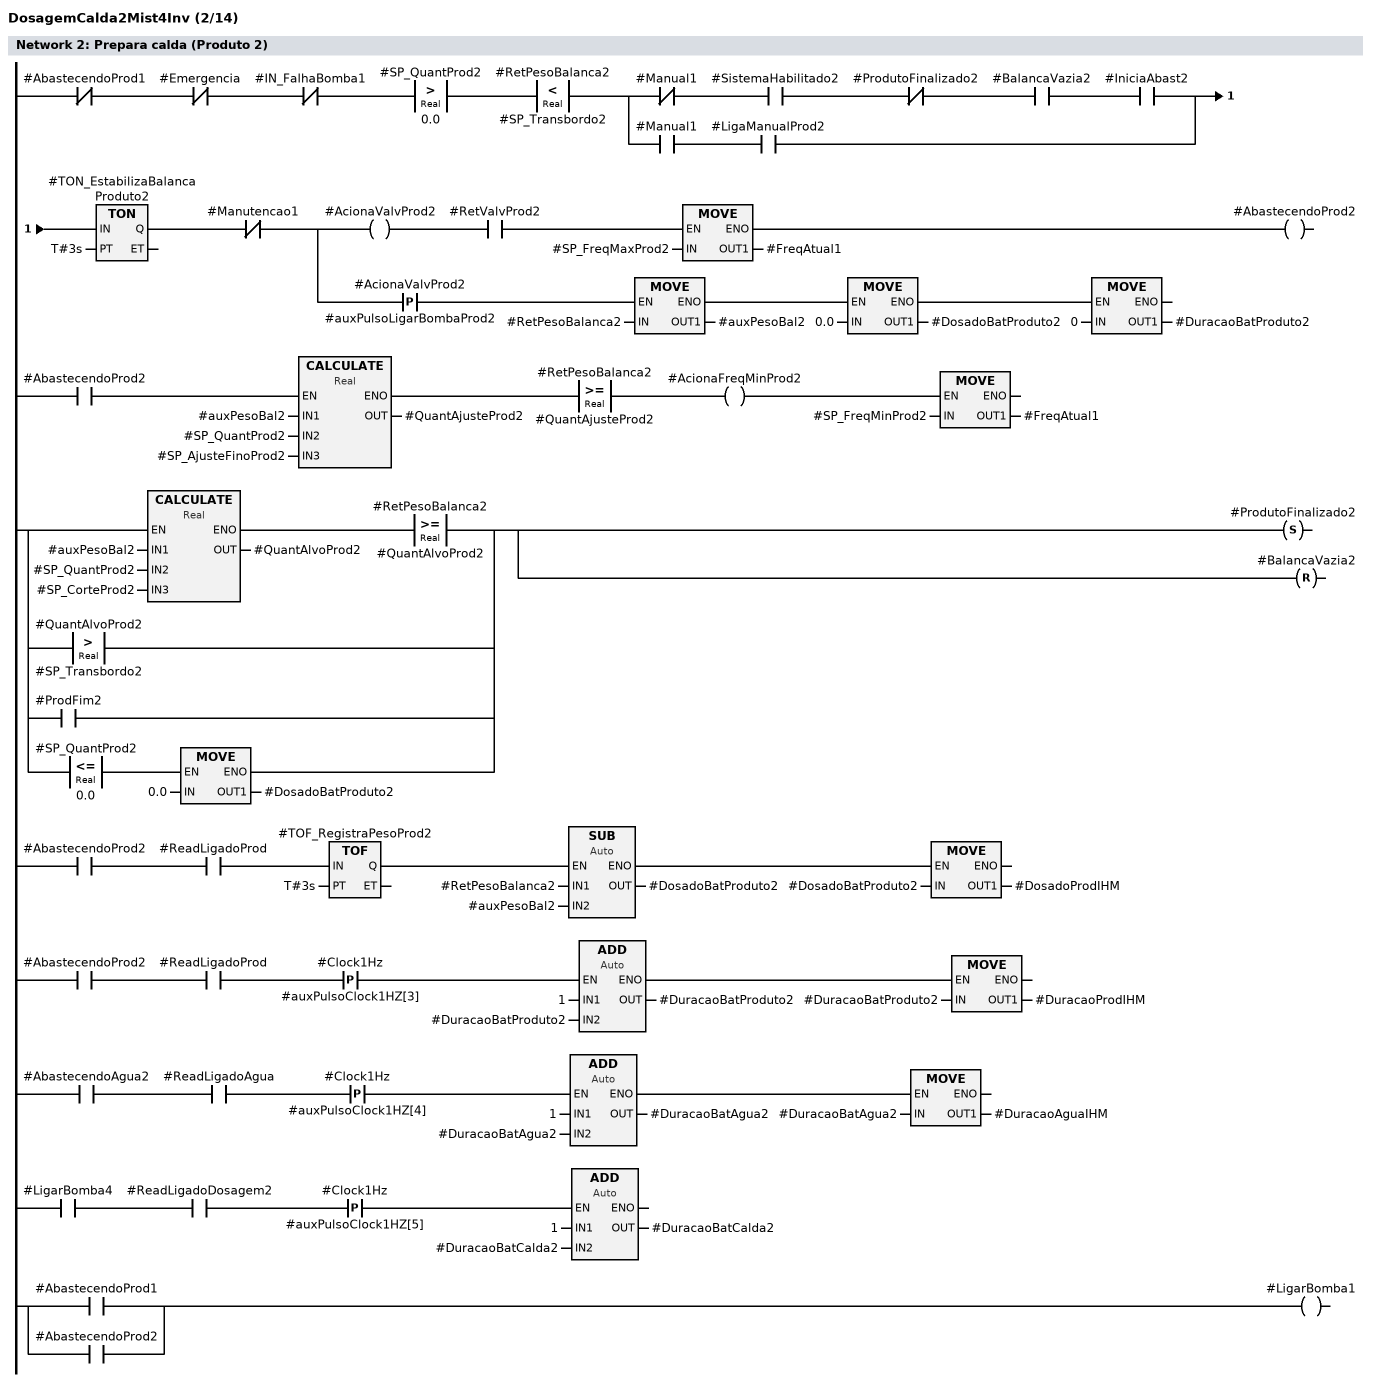
   #TON_EstabilizaBalancaProduto2(IN := NOT #AbastecendoProd1 AND NOT #Emergencia AND NOT #IN_FalhaBomba1 AND (#SP_QuantProd2 > 0.0) AND (#RetPesoBalanca2 < #SP_Transbordo2) AND ((NOT #Manual1 AND #SistemaHabilitado2 AND NOT #ProdutoFinalizado2 AND #BalancaVazia2 AND #IniciaAbast2) OR (#Manual1 AND #LigaManualProd2)),   // TON
                           PT := T#3s);
   #AcionaValvProd2 := #TON_EstabilizaBalancaProduto2.Q AND NOT #Manutencao1;
   #_w1 := #AcionaValvProd2 AND #RetValvProd2;
   IF #_w1 THEN #FreqAtual1 := #SP_FreqMaxProd2; END_IF;
   #AbastecendoProd2 := #_w1;
   #_w2 := #AcionaValvProd2 AND #AcionaValvProd2 AND NOT #auxPulsoLigarBombaProd2;   // rising edge of #AcionaValvProd2
   #auxPulsoLigarBombaProd2 := #AcionaValvProd2;
   IF #_w2 THEN
       #auxPesoBal2 := #RetPesoBalanca2;
       #DosadoBatProduto2 := 0.0;
       #DuracaoBatProduto2 := 0;
   END_IF;
   IF #AbastecendoProd2 THEN
       #QuantAjusteProd2 := (#auxPesoBal2 + #SP_QuantProd2 - #SP_AjusteFinoProd2);
   END_IF;
   #AcionaFreqMinProd2 := #AbastecendoProd2 AND (#RetPesoBalanca2 >= #QuantAjusteProd2);
   IF #AcionaFreqMinProd2 THEN #FreqAtual1 := #SP_FreqMinProd2; END_IF;
   #QuantAlvoProd2 := (#auxPesoBal2 + #SP_QuantProd2 - #SP_CorteProd2);
   #_w3 := #SP_QuantProd2 <= 0.0;
   IF #_w3 THEN #DosadoBatProduto2 := 0.0; END_IF;
   IF (#RetPesoBalanca2 >= #QuantAlvoProd2) OR (#QuantAlvoProd2 > #SP_Transbordo2) OR #ProdFim2 OR #_w3 THEN
       #ProdutoFinalizado2 := TRUE;
       #BalancaVazia2 := FALSE;
   END_IF;
   #TOF_RegistraPesoProd2(IN := #AbastecendoProd2 AND #ReadLigadoProd, PT := T#3s);   // TOF
   IF #TOF_RegistraPesoProd2.Q THEN
       #DosadoBatProduto2 := #RetPesoBalanca2 - #auxPesoBal2;
       #DosadoProdIHM := #DosadoBatProduto2;
   END_IF;
   #_w4 := #AbastecendoProd2 AND #ReadLigadoProd AND #Clock1Hz AND NOT #auxPulsoClock1HZ[3];   // rising edge of #Clock1Hz
   #auxPulsoClock1HZ[3] := #Clock1Hz;
   IF #_w4 THEN
       #DuracaoBatProduto2 := 1 + #DuracaoBatProduto2;
       #DuracaoProdIHM := #DuracaoBatProduto2;
   END_IF;
   #_w5 := #AbastecendoAgua2 AND #ReadLigadoAgua AND #Clock1Hz AND NOT #auxPulsoClock1HZ[4];   // rising edge of #Clock1Hz
   #auxPulsoClock1HZ[4] := #Clock1Hz;
   IF #_w5 THEN
       #DuracaoBatAgua2 := 1 + #DuracaoBatAgua2;
       #DuracaoAguaIHM := #DuracaoBatAgua2;
   END_IF;
   #_w6 := #LigarBomba4 AND #ReadLigadoDosagem2 AND #Clock1Hz AND NOT #auxPulsoClock1HZ[5];   // rising edge of #Clock1Hz
   #auxPulsoClock1HZ[5] := #Clock1Hz;
   IF #_w6 THEN #DuracaoBatCalda2 := 1 + #DuracaoBatCalda2; END_IF;
   #LigarBomba1 := #AbastecendoProd1 OR #AbastecendoProd2;
END_REGION

REGION Network 3: Prepara calda (Agua 1)
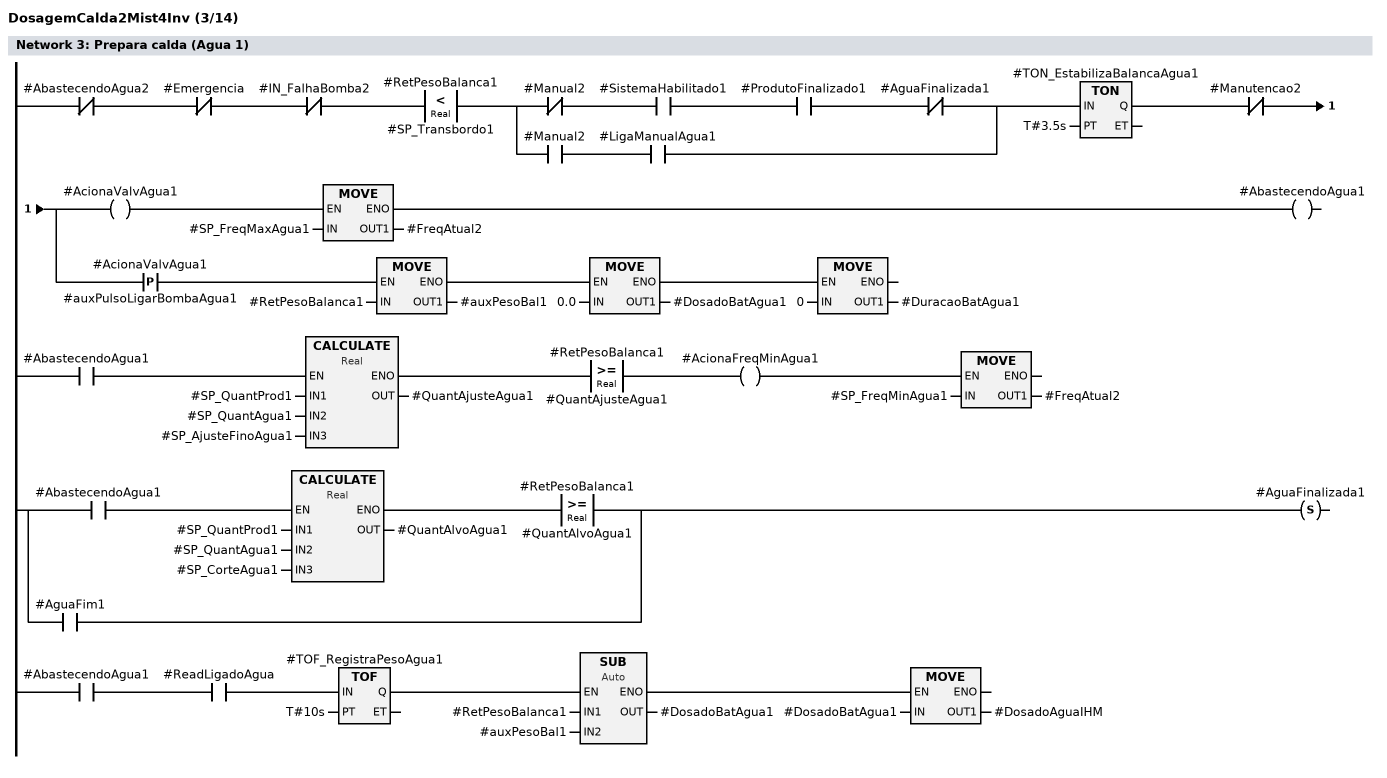
   #TON_EstabilizaBalancaAgua1(IN := NOT #AbastecendoAgua2 AND NOT #Emergencia AND NOT #IN_FalhaBomba2 AND (#RetPesoBalanca1 < #SP_Transbordo1) AND ((NOT #Manual2 AND #SistemaHabilitado1 AND #ProdutoFinalizado1 AND NOT #AguaFinalizada1) OR (#Manual2 AND #LigaManualAgua1)),   // TON
                           PT := T#3.5s);
   #AcionaValvAgua1 := #TON_EstabilizaBalancaAgua1.Q AND NOT #Manutencao2;
   IF #AcionaValvAgua1 THEN #FreqAtual2 := #SP_FreqMaxAgua1; END_IF;
   #AbastecendoAgua1 := #AcionaValvAgua1;
   #_w1 := #AcionaValvAgua1 AND #AcionaValvAgua1 AND NOT #auxPulsoLigarBombaAgua1;   // rising edge of #AcionaValvAgua1
   #auxPulsoLigarBombaAgua1 := #AcionaValvAgua1;
   IF #_w1 THEN
       #auxPesoBal1 := #RetPesoBalanca1;
       #DosadoBatAgua1 := 0.0;
       #DuracaoBatAgua1 := 0;
   END_IF;
   IF #AbastecendoAgua1 THEN
       #QuantAjusteAgua1 := (#SP_QuantProd1 + #SP_QuantAgua1 - #SP_AjusteFinoAgua1);
   END_IF;
   #AcionaFreqMinAgua1 := #AbastecendoAgua1 AND (#RetPesoBalanca1 >= #QuantAjusteAgua1);
   IF #AcionaFreqMinAgua1 THEN #FreqAtual2 := #SP_FreqMinAgua1; END_IF;
   IF #AbastecendoAgua1 THEN #QuantAlvoAgua1 := (#SP_QuantProd1 + #SP_QuantAgua1 - #SP_CorteAgua1); END_IF;
   IF (#AbastecendoAgua1 AND (#RetPesoBalanca1 >= #QuantAlvoAgua1)) OR #AguaFim1 THEN
       #AguaFinalizada1 := TRUE;
   END_IF;
   #TOF_RegistraPesoAgua1(IN := #AbastecendoAgua1 AND #ReadLigadoAgua, PT := T#10s);   // TOF
   IF #TOF_RegistraPesoAgua1.Q THEN
       #DosadoBatAgua1 := #RetPesoBalanca1 - #auxPesoBal1;
       #DosadoAguaIHM := #DosadoBatAgua1;
   END_IF;
END_REGION

REGION Network 4: Prepara calda (Agua 2)
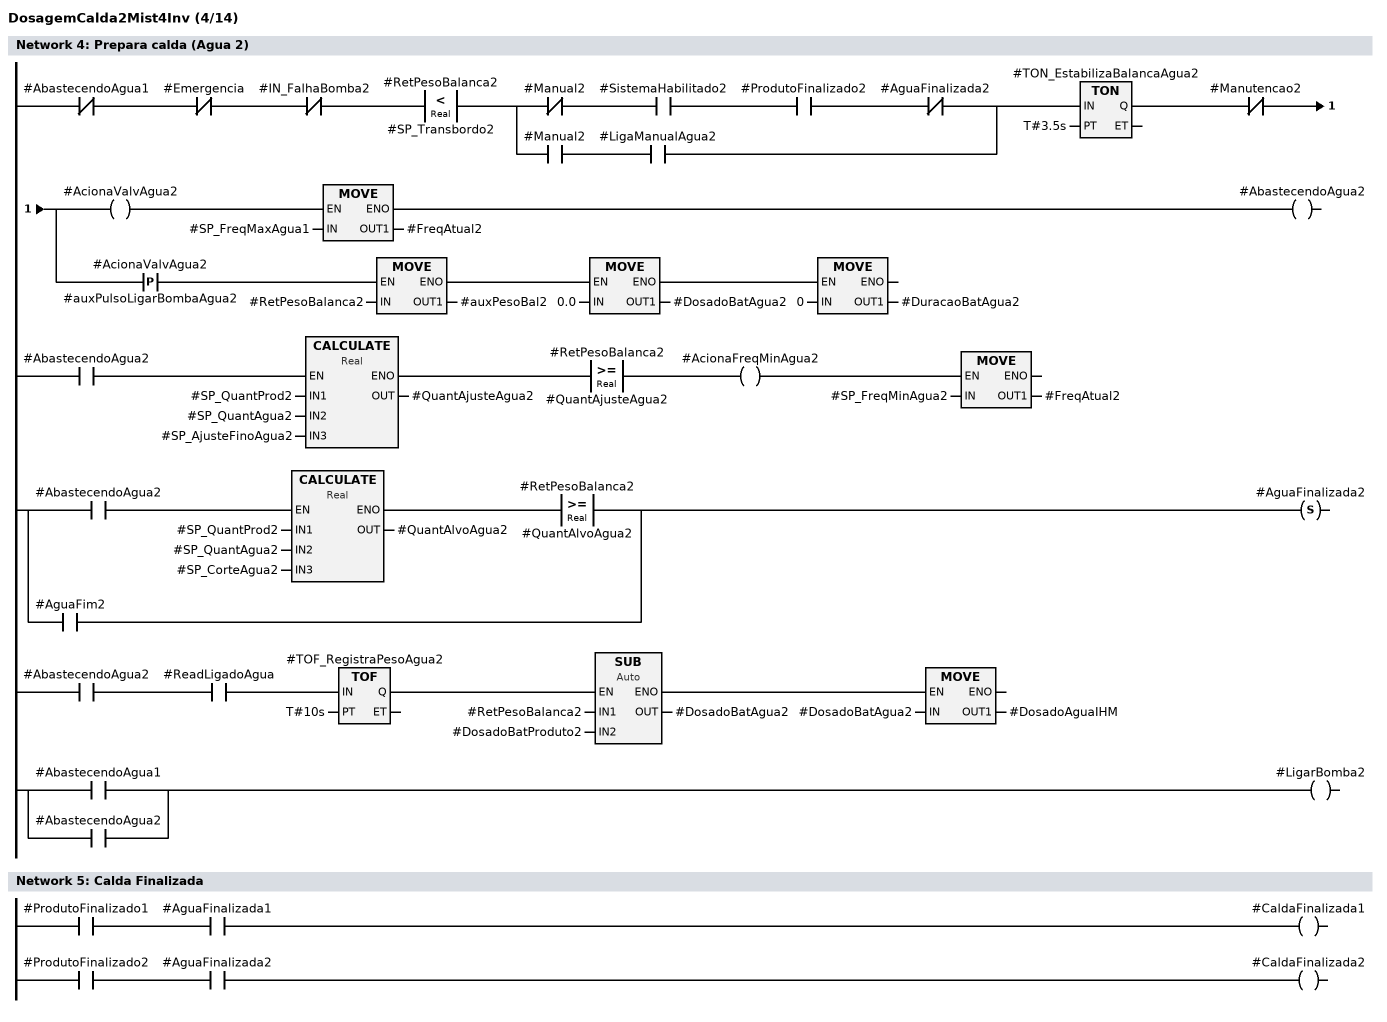
   #TON_EstabilizaBalancaAgua2(IN := NOT #AbastecendoAgua1 AND NOT #Emergencia AND NOT #IN_FalhaBomba2 AND (#RetPesoBalanca2 < #SP_Transbordo2) AND ((NOT #Manual2 AND #SistemaHabilitado2 AND #ProdutoFinalizado2 AND NOT #AguaFinalizada2) OR (#Manual2 AND #LigaManualAgua2)),   // TON
                           PT := T#3.5s);
   #AcionaValvAgua2 := #TON_EstabilizaBalancaAgua2.Q AND NOT #Manutencao2;
   IF #AcionaValvAgua2 THEN #FreqAtual2 := #SP_FreqMaxAgua1; END_IF;
   #AbastecendoAgua2 := #AcionaValvAgua2;
   #_w1 := #AcionaValvAgua2 AND #AcionaValvAgua2 AND NOT #auxPulsoLigarBombaAgua2;   // rising edge of #AcionaValvAgua2
   #auxPulsoLigarBombaAgua2 := #AcionaValvAgua2;
   IF #_w1 THEN
       #auxPesoBal2 := #RetPesoBalanca2;
       #DosadoBatAgua2 := 0.0;
       #DuracaoBatAgua2 := 0;
   END_IF;
   IF #AbastecendoAgua2 THEN
       #QuantAjusteAgua2 := (#SP_QuantProd2 + #SP_QuantAgua2 - #SP_AjusteFinoAgua2);
   END_IF;
   #AcionaFreqMinAgua2 := #AbastecendoAgua2 AND (#RetPesoBalanca2 >= #QuantAjusteAgua2);
   IF #AcionaFreqMinAgua2 THEN #FreqAtual2 := #SP_FreqMinAgua2; END_IF;
   IF #AbastecendoAgua2 THEN #QuantAlvoAgua2 := (#SP_QuantProd2 + #SP_QuantAgua2 - #SP_CorteAgua2); END_IF;
   IF (#AbastecendoAgua2 AND (#RetPesoBalanca2 >= #QuantAlvoAgua2)) OR #AguaFim2 THEN
       #AguaFinalizada2 := TRUE;
   END_IF;
   #TOF_RegistraPesoAgua2(IN := #AbastecendoAgua2 AND #ReadLigadoAgua, PT := T#10s);   // TOF
   IF #TOF_RegistraPesoAgua2.Q THEN
       #DosadoBatAgua2 := #RetPesoBalanca2 - #DosadoBatProduto2;
       #DosadoAguaIHM := #DosadoBatAgua2;
   END_IF;
   #LigarBomba2 := #AbastecendoAgua1 OR #AbastecendoAgua2;
END_REGION

REGION Network 5: Calda Finalizada
   RUNG wire#powerrail
      Contact( #ProdutoFinalizado1 )
      Contact( #AguaFinalizada1 )
      Coil( #CaldaFinalizada1 )
   END_RUNG
   RUNG wire#powerrail
      Contact( #ProdutoFinalizado2 )
      Contact( #AguaFinalizada2 )
      Coil( #CaldaFinalizada2 )
   END_RUNG
   // the same network as SCL:
   #CaldaFinalizada1 := #ProdutoFinalizado1 AND #AguaFinalizada1;
   #CaldaFinalizada2 := #ProdutoFinalizado2 AND #AguaFinalizada2;
END_REGION

REGION Network 6: Tempo de mistura seca 1
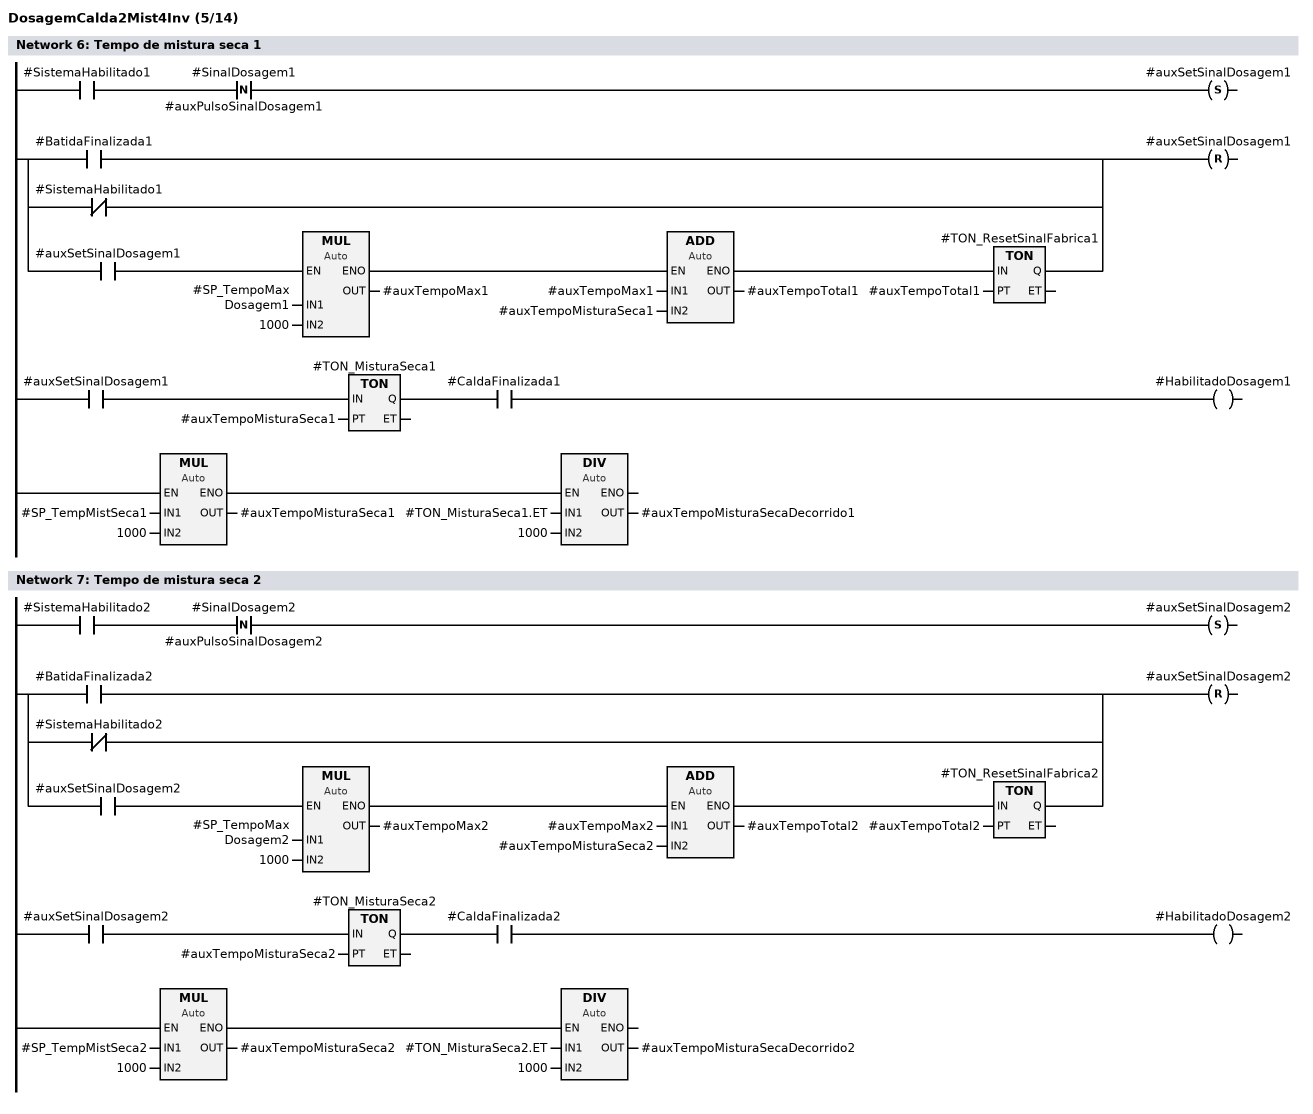
   #_w1 := #SistemaHabilitado1 AND NOT #SinalDosagem1 AND #auxPulsoSinalDosagem1;   // falling edge of #SinalDosagem1
   #auxPulsoSinalDosagem1 := #SinalDosagem1;
   IF #_w1 THEN #auxSetSinalDosagem1 := TRUE; END_IF;
   IF #auxSetSinalDosagem1 THEN
       #auxTempoMax1 := #SP_TempoMaxDosagem1 * 1000;
       #auxTempoTotal1 := #auxTempoMax1 + #auxTempoMisturaSeca1;
   END_IF;
   #TON_ResetSinalFabrica1(IN := #auxSetSinalDosagem1, PT := #auxTempoTotal1);   // TON
   IF #BatidaFinalizada1 OR NOT #SistemaHabilitado1 OR #TON_ResetSinalFabrica1.Q THEN
       #auxSetSinalDosagem1 := FALSE;
   END_IF;
   #TON_MisturaSeca1(IN := #auxSetSinalDosagem1, PT := #auxTempoMisturaSeca1);   // TON
   #HabilitadoDosagem1 := #TON_MisturaSeca1.Q AND #CaldaFinalizada1;
   #auxTempoMisturaSeca1 := #SP_TempMistSeca1 * 1000;
   #auxTempoMisturaSecaDecorrido1 := #TON_MisturaSeca1.ET / 1000;
END_REGION

REGION Network 7: Tempo de mistura seca 2
   #_w1 := #SistemaHabilitado2 AND NOT #SinalDosagem2 AND #auxPulsoSinalDosagem2;   // falling edge of #SinalDosagem2
   #auxPulsoSinalDosagem2 := #SinalDosagem2;
   IF #_w1 THEN #auxSetSinalDosagem2 := TRUE; END_IF;
   IF #auxSetSinalDosagem2 THEN
       #auxTempoMax2 := #SP_TempoMaxDosagem2 * 1000;
       #auxTempoTotal2 := #auxTempoMax2 + #auxTempoMisturaSeca2;
   END_IF;
   #TON_ResetSinalFabrica2(IN := #auxSetSinalDosagem2, PT := #auxTempoTotal2);   // TON
   IF #BatidaFinalizada2 OR NOT #SistemaHabilitado2 OR #TON_ResetSinalFabrica2.Q THEN
       #auxSetSinalDosagem2 := FALSE;
   END_IF;
   #TON_MisturaSeca2(IN := #auxSetSinalDosagem2, PT := #auxTempoMisturaSeca2);   // TON
   #HabilitadoDosagem2 := #TON_MisturaSeca2.Q AND #CaldaFinalizada2;
   #auxTempoMisturaSeca2 := #SP_TempMistSeca2 * 1000;
   #auxTempoMisturaSecaDecorrido2 := #TON_MisturaSeca2.ET / 1000;
END_REGION

REGION Network 8: Dosa calda 1
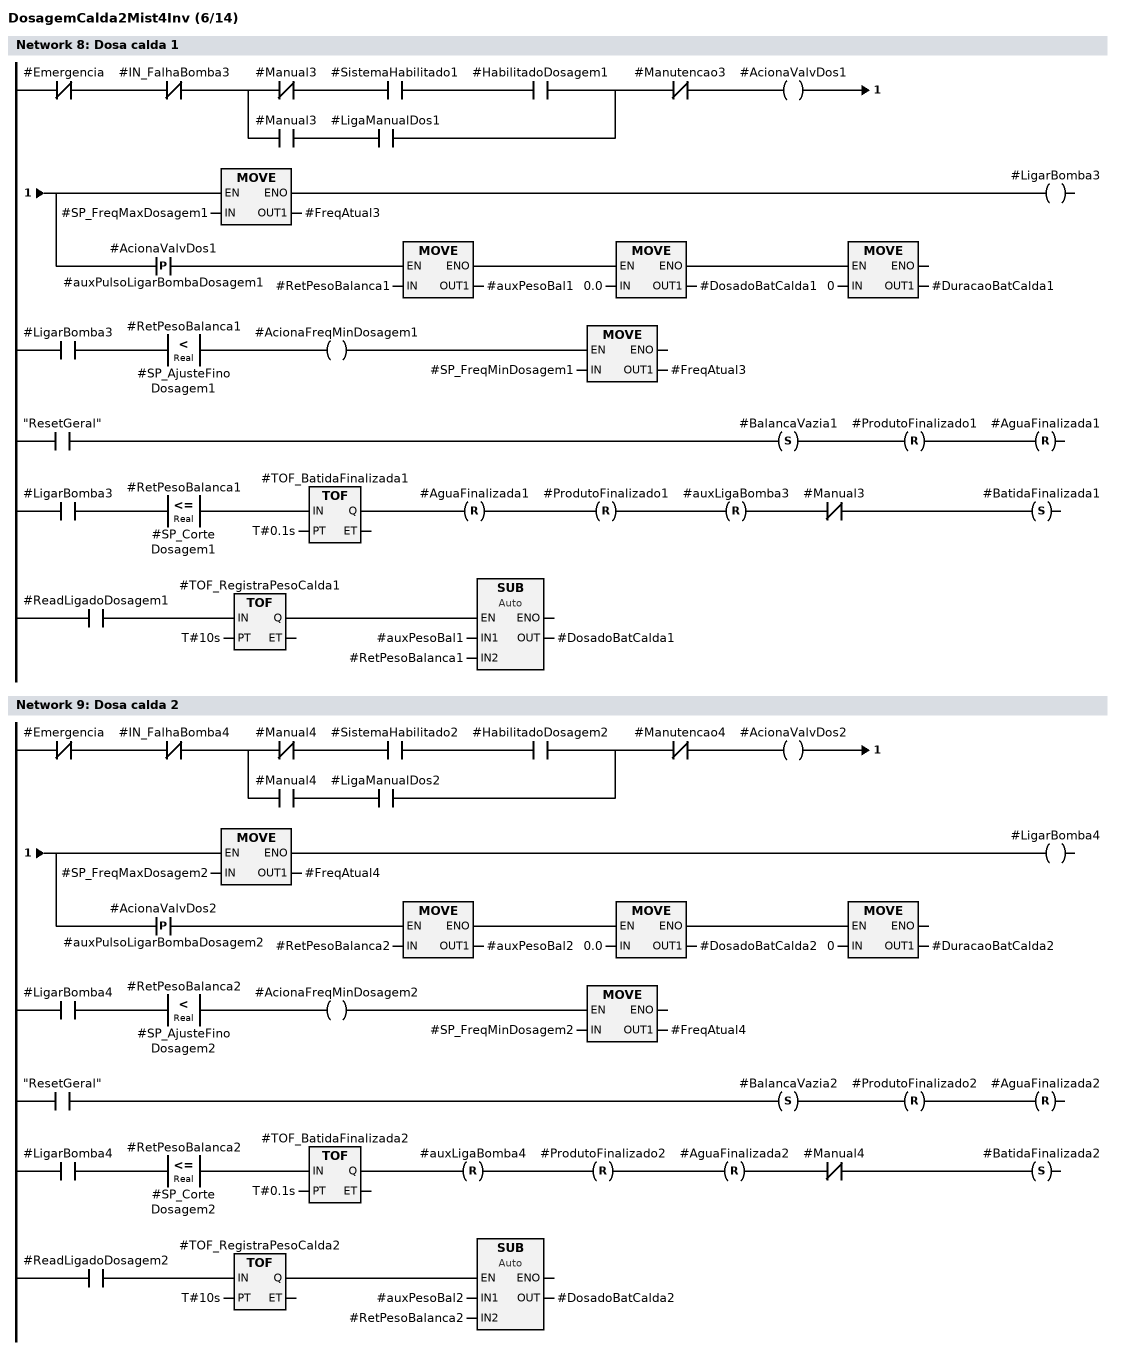
   #AcionaValvDos1 := NOT #Emergencia AND NOT #IN_FalhaBomba3 AND ((NOT #Manual3 AND #SistemaHabilitado1 AND #HabilitadoDosagem1) OR (#Manual3 AND #LigaManualDos1)) AND NOT #Manutencao3;
   IF #AcionaValvDos1 THEN #FreqAtual3 := #SP_FreqMaxDosagem1; END_IF;
   #LigarBomba3 := #AcionaValvDos1;
   #_w1 := #AcionaValvDos1 AND #AcionaValvDos1 AND NOT #auxPulsoLigarBombaDosagem1;   // rising edge of #AcionaValvDos1
   #auxPulsoLigarBombaDosagem1 := #AcionaValvDos1;
   IF #_w1 THEN
       #auxPesoBal1 := #RetPesoBalanca1;
       #DosadoBatCalda1 := 0.0;
       #DuracaoBatCalda1 := 0;
   END_IF;
   #AcionaFreqMinDosagem1 := #LigarBomba3 AND (#RetPesoBalanca1 < #SP_AjusteFinoDosagem1);
   IF #AcionaFreqMinDosagem1 THEN #FreqAtual3 := #SP_FreqMinDosagem1; END_IF;
   IF "ResetGeral" THEN
       #BalancaVazia1 := TRUE;
       #ProdutoFinalizado1 := FALSE;
       #AguaFinalizada1 := FALSE;
   END_IF;
   #TOF_BatidaFinalizada1(IN := #LigarBomba3 AND (#RetPesoBalanca1 <= #SP_CorteDosagem1), PT := T#0.1s);   // TOF
   IF #TOF_BatidaFinalizada1.Q THEN
       #AguaFinalizada1 := FALSE;
       #ProdutoFinalizado1 := FALSE;
       #auxLigaBomba3 := FALSE;
   END_IF;
   IF #TOF_BatidaFinalizada1.Q AND NOT #Manual3 THEN #BatidaFinalizada1 := TRUE; END_IF;
   #TOF_RegistraPesoCalda1(IN := #ReadLigadoDosagem1, PT := T#10s);   // TOF
   IF #TOF_RegistraPesoCalda1.Q THEN #DosadoBatCalda1 := #auxPesoBal1 - #RetPesoBalanca1; END_IF;
END_REGION

REGION Network 9: Dosa calda 2
   #AcionaValvDos2 := NOT #Emergencia AND NOT #IN_FalhaBomba4 AND ((NOT #Manual4 AND #SistemaHabilitado2 AND #HabilitadoDosagem2) OR (#Manual4 AND #LigaManualDos2)) AND NOT #Manutencao4;
   IF #AcionaValvDos2 THEN #FreqAtual4 := #SP_FreqMaxDosagem2; END_IF;
   #LigarBomba4 := #AcionaValvDos2;
   #_w1 := #AcionaValvDos2 AND #AcionaValvDos2 AND NOT #auxPulsoLigarBombaDosagem2;   // rising edge of #AcionaValvDos2
   #auxPulsoLigarBombaDosagem2 := #AcionaValvDos2;
   IF #_w1 THEN
       #auxPesoBal2 := #RetPesoBalanca2;
       #DosadoBatCalda2 := 0.0;
       #DuracaoBatCalda2 := 0;
   END_IF;
   #AcionaFreqMinDosagem2 := #LigarBomba4 AND (#RetPesoBalanca2 < #SP_AjusteFinoDosagem2);
   IF #AcionaFreqMinDosagem2 THEN #FreqAtual4 := #SP_FreqMinDosagem2; END_IF;
   IF "ResetGeral" THEN
       #BalancaVazia2 := TRUE;
       #ProdutoFinalizado2 := FALSE;
       #AguaFinalizada2 := FALSE;
   END_IF;
   #TOF_BatidaFinalizada2(IN := #LigarBomba4 AND (#RetPesoBalanca2 <= #SP_CorteDosagem2), PT := T#0.1s);   // TOF
   IF #TOF_BatidaFinalizada2.Q THEN
       #auxLigaBomba4 := FALSE;
       #ProdutoFinalizado2 := FALSE;
       #AguaFinalizada2 := FALSE;
   END_IF;
   IF #TOF_BatidaFinalizada2.Q AND NOT #Manual4 THEN #BatidaFinalizada2 := TRUE; END_IF;
   #TOF_RegistraPesoCalda2(IN := #ReadLigadoDosagem2, PT := T#10s);   // TOF
   IF #TOF_RegistraPesoCalda2.Q THEN #DosadoBatCalda2 := #auxPesoBal2 - #RetPesoBalanca2; END_IF;
END_REGION

REGION Network 10: Grava batelada
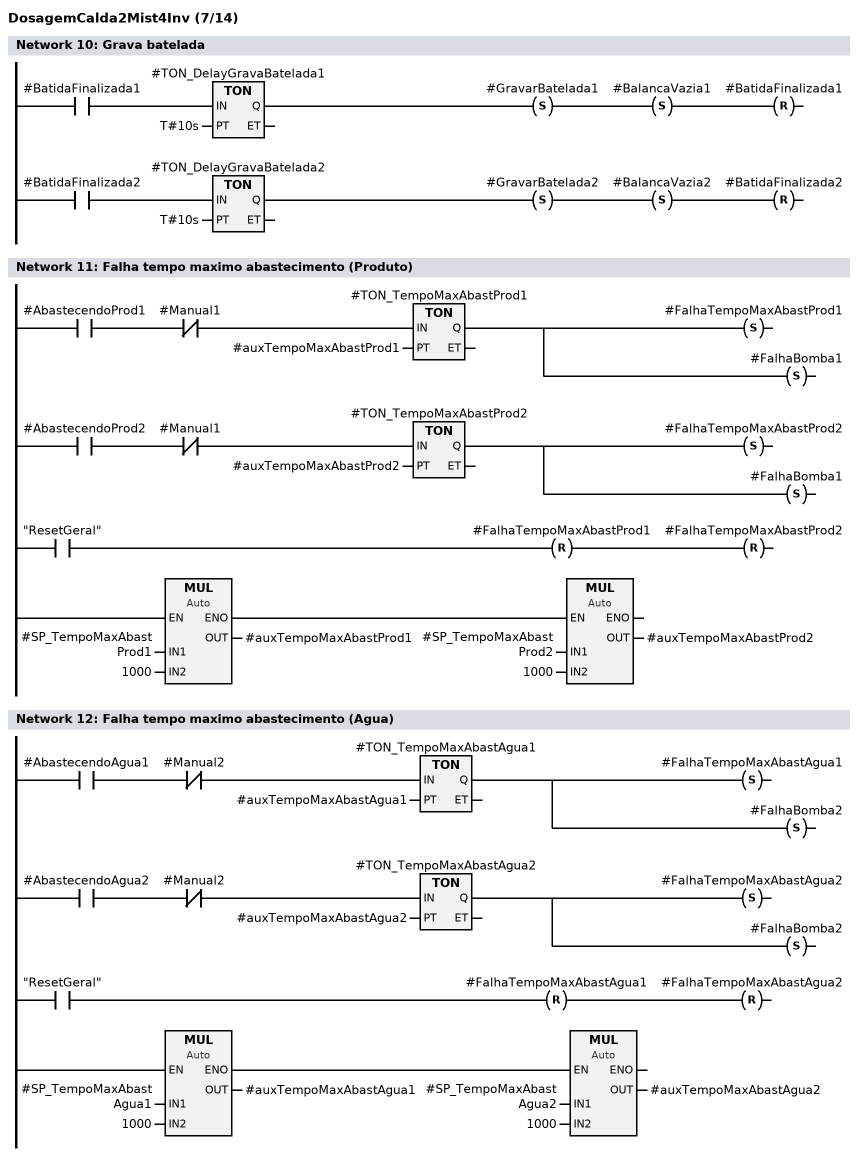
   #TON_DelayGravaBatelada1(IN := #BatidaFinalizada1, PT := T#10s);   // TON
   IF #TON_DelayGravaBatelada1.Q THEN
       #GravarBatelada1 := TRUE;
       #BalancaVazia1 := TRUE;
       #BatidaFinalizada1 := FALSE;
   END_IF;
   #TON_DelayGravaBatelada2(IN := #BatidaFinalizada2, PT := T#10s);   // TON
   IF #TON_DelayGravaBatelada2.Q THEN
       #GravarBatelada2 := TRUE;
       #BalancaVazia2 := TRUE;
       #BatidaFinalizada2 := FALSE;
   END_IF;
END_REGION

REGION Network 11: Falha tempo maximo abastecimento (Produto)
   #TON_TempoMaxAbastProd1(IN := #AbastecendoProd1 AND NOT #Manual1, PT := #auxTempoMaxAbastProd1);   // TON
   IF #TON_TempoMaxAbastProd1.Q THEN
       #FalhaTempoMaxAbastProd1 := TRUE;
       #FalhaBomba1 := TRUE;
   END_IF;
   #TON_TempoMaxAbastProd2(IN := #AbastecendoProd2 AND NOT #Manual1, PT := #auxTempoMaxAbastProd2);   // TON
   IF #TON_TempoMaxAbastProd2.Q THEN
       #FalhaTempoMaxAbastProd2 := TRUE;
       #FalhaBomba1 := TRUE;
   END_IF;
   IF "ResetGeral" THEN
       #FalhaTempoMaxAbastProd1 := FALSE;
       #FalhaTempoMaxAbastProd2 := FALSE;
   END_IF;
   #auxTempoMaxAbastProd1 := #SP_TempoMaxAbastProd1 * 1000;
   #auxTempoMaxAbastProd2 := #SP_TempoMaxAbastProd2 * 1000;
END_REGION

REGION Network 12: Falha tempo maximo abastecimento (Agua)
   #TON_TempoMaxAbastAgua1(IN := #AbastecendoAgua1 AND NOT #Manual2, PT := #auxTempoMaxAbastAgua1);   // TON
   IF #TON_TempoMaxAbastAgua1.Q THEN
       #FalhaTempoMaxAbastAgua1 := TRUE;
       #FalhaBomba2 := TRUE;
   END_IF;
   #TON_TempoMaxAbastAgua2(IN := #AbastecendoAgua2 AND NOT #Manual2, PT := #auxTempoMaxAbastAgua2);   // TON
   IF #TON_TempoMaxAbastAgua2.Q THEN
       #FalhaTempoMaxAbastAgua2 := TRUE;
       #FalhaBomba2 := TRUE;
   END_IF;
   IF "ResetGeral" THEN
       #FalhaTempoMaxAbastAgua1 := FALSE;
       #FalhaTempoMaxAbastAgua2 := FALSE;
   END_IF;
   #auxTempoMaxAbastAgua1 := #SP_TempoMaxAbastAgua1 * 1000;
   #auxTempoMaxAbastAgua2 := #SP_TempoMaxAbastAgua2 * 1000;
END_REGION

REGION Network 13: Falha tempo maximo de dosagem (Calda)
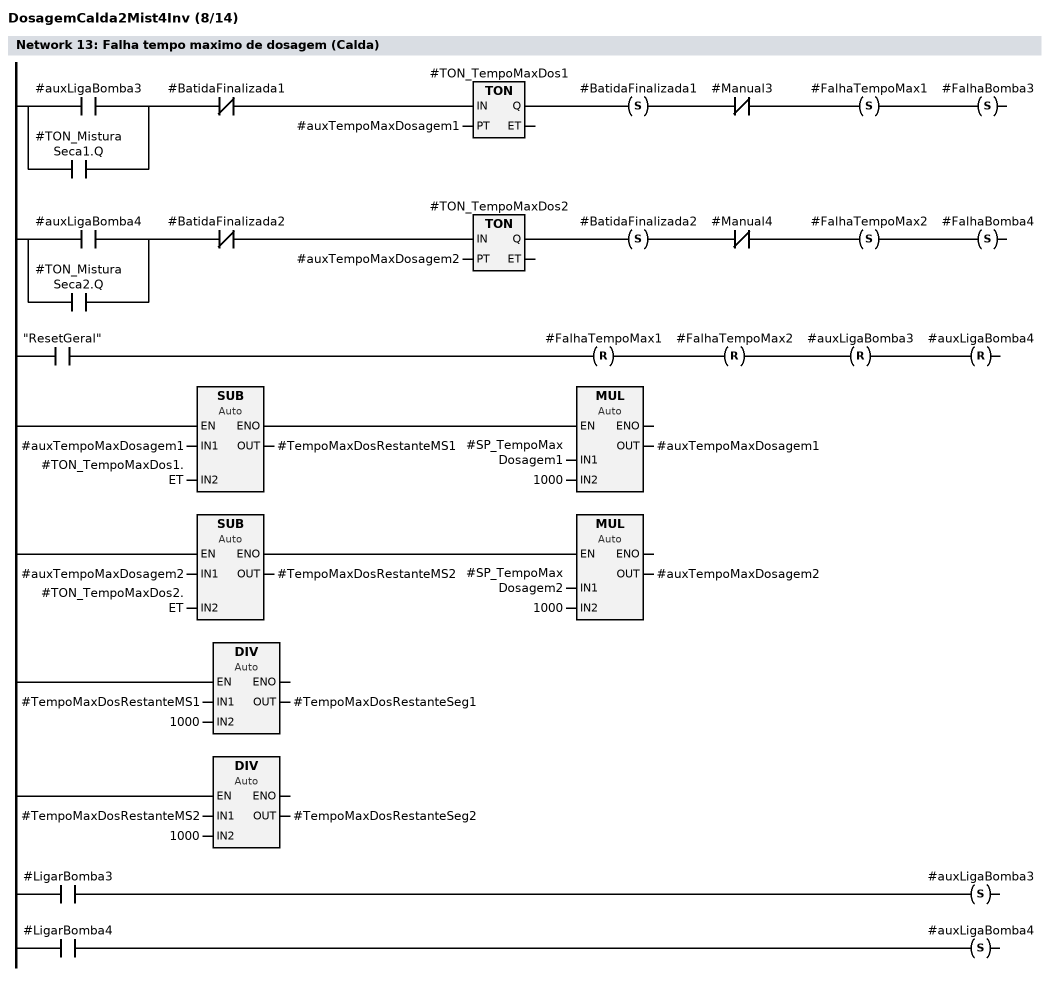
   #TON_TempoMaxDos1(IN := (#auxLigaBomba3 OR #TON_MisturaSeca1.Q) AND NOT #BatidaFinalizada1,   // TON
                     PT := #auxTempoMaxDosagem1);
   IF #TON_TempoMaxDos1.Q THEN #BatidaFinalizada1 := TRUE; END_IF;
   IF #TON_TempoMaxDos1.Q AND NOT #Manual3 THEN
       #FalhaTempoMax1 := TRUE;
       #FalhaBomba3 := TRUE;
   END_IF;
   #TON_TempoMaxDos2(IN := (#auxLigaBomba4 OR #TON_MisturaSeca2.Q) AND NOT #BatidaFinalizada2,   // TON
                     PT := #auxTempoMaxDosagem2);
   IF #TON_TempoMaxDos2.Q THEN #BatidaFinalizada2 := TRUE; END_IF;
   IF #TON_TempoMaxDos2.Q AND NOT #Manual4 THEN
       #FalhaTempoMax2 := TRUE;
       #FalhaBomba4 := TRUE;
   END_IF;
   IF "ResetGeral" THEN
       #FalhaTempoMax1 := FALSE;
       #FalhaTempoMax2 := FALSE;
       #auxLigaBomba3 := FALSE;
       #auxLigaBomba4 := FALSE;
   END_IF;
   #TempoMaxDosRestanteMS1 := #auxTempoMaxDosagem1 - #TON_TempoMaxDos1.ET;
   #auxTempoMaxDosagem1 := #SP_TempoMaxDosagem1 * 1000;
   #TempoMaxDosRestanteMS2 := #auxTempoMaxDosagem2 - #TON_TempoMaxDos2.ET;
   #auxTempoMaxDosagem2 := #SP_TempoMaxDosagem2 * 1000;
   #TempoMaxDosRestanteSeg1 := #TempoMaxDosRestanteMS1 / 1000;
   #TempoMaxDosRestanteSeg2 := #TempoMaxDosRestanteMS2 / 1000;
   IF #LigarBomba3 THEN #auxLigaBomba3 := TRUE; END_IF;
   IF #LigarBomba4 THEN #auxLigaBomba4 := TRUE; END_IF;
END_REGION

REGION Network 14: Falha bombas
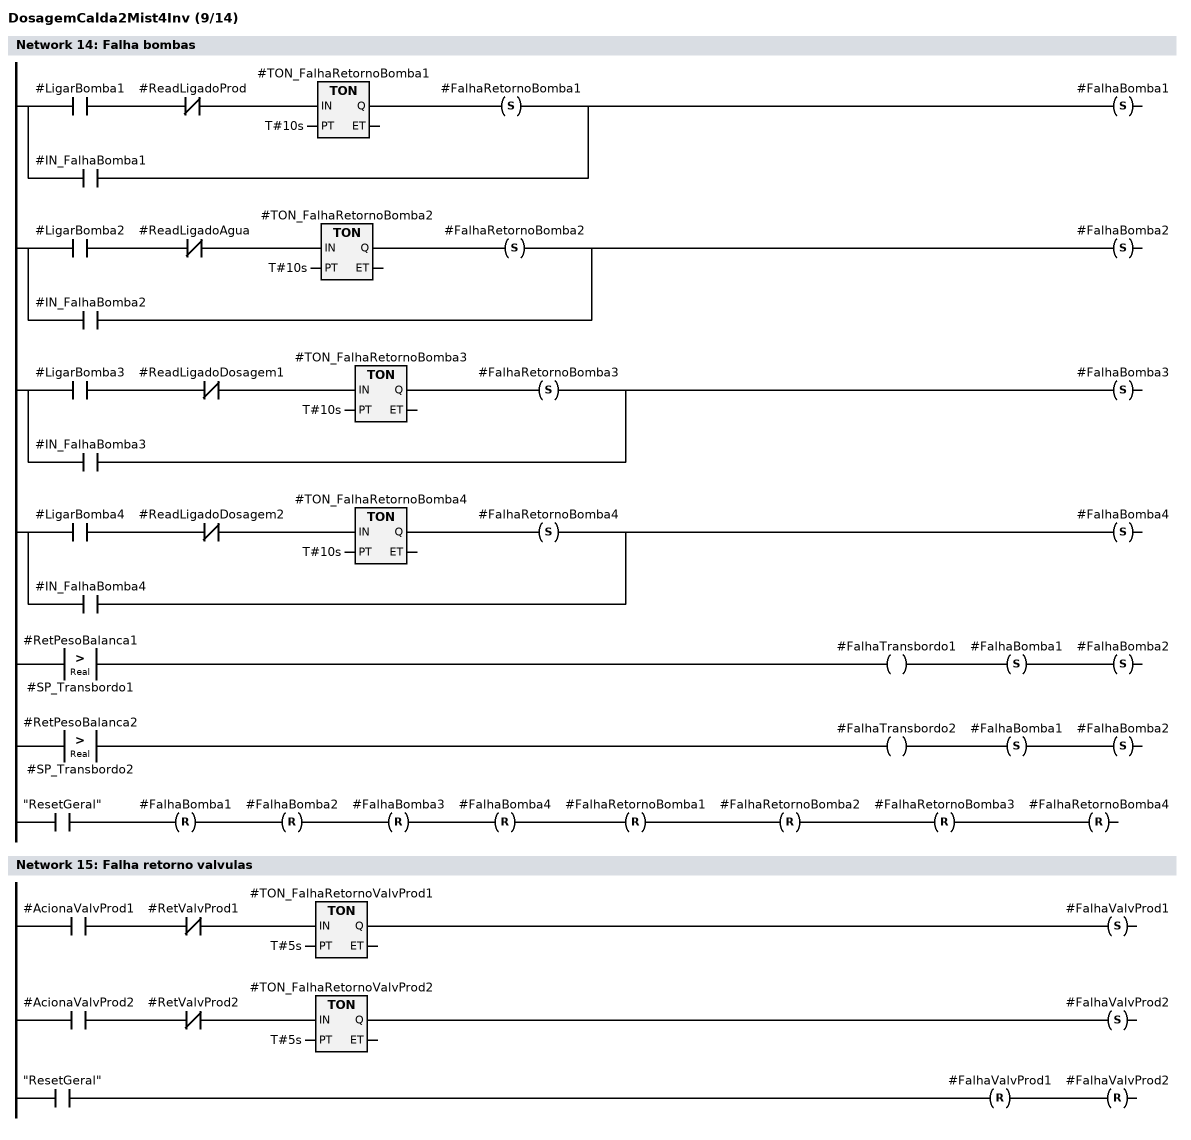
   #TON_FalhaRetornoBomba1(IN := #LigarBomba1 AND NOT #ReadLigadoProd, PT := T#10s);   // TON
   IF #TON_FalhaRetornoBomba1.Q THEN #FalhaRetornoBomba1 := TRUE; END_IF;
   IF #TON_FalhaRetornoBomba1.Q OR #IN_FalhaBomba1 THEN #FalhaBomba1 := TRUE; END_IF;
   #TON_FalhaRetornoBomba2(IN := #LigarBomba2 AND NOT #ReadLigadoAgua, PT := T#10s);   // TON
   IF #TON_FalhaRetornoBomba2.Q THEN #FalhaRetornoBomba2 := TRUE; END_IF;
   IF #TON_FalhaRetornoBomba2.Q OR #IN_FalhaBomba2 THEN #FalhaBomba2 := TRUE; END_IF;
   #TON_FalhaRetornoBomba3(IN := #LigarBomba3 AND NOT #ReadLigadoDosagem1, PT := T#10s);   // TON
   IF #TON_FalhaRetornoBomba3.Q THEN #FalhaRetornoBomba3 := TRUE; END_IF;
   IF #TON_FalhaRetornoBomba3.Q OR #IN_FalhaBomba3 THEN #FalhaBomba3 := TRUE; END_IF;
   #TON_FalhaRetornoBomba4(IN := #LigarBomba4 AND NOT #ReadLigadoDosagem2, PT := T#10s);   // TON
   IF #TON_FalhaRetornoBomba4.Q THEN #FalhaRetornoBomba4 := TRUE; END_IF;
   IF #TON_FalhaRetornoBomba4.Q OR #IN_FalhaBomba4 THEN #FalhaBomba4 := TRUE; END_IF;
   #FalhaTransbordo1 := #RetPesoBalanca1 > #SP_Transbordo1;
   IF #FalhaTransbordo1 THEN
       #FalhaBomba1 := TRUE;
       #FalhaBomba2 := TRUE;
   END_IF;
   #FalhaTransbordo2 := #RetPesoBalanca2 > #SP_Transbordo2;
   IF #FalhaTransbordo2 THEN
       #FalhaBomba1 := TRUE;
       #FalhaBomba2 := TRUE;
   END_IF;
   IF "ResetGeral" THEN
       #FalhaBomba1 := FALSE;
       #FalhaBomba2 := FALSE;
       #FalhaBomba3 := FALSE;
       #FalhaBomba4 := FALSE;
       #FalhaRetornoBomba1 := FALSE;
       #FalhaRetornoBomba2 := FALSE;
       #FalhaRetornoBomba3 := FALSE;
       #FalhaRetornoBomba4 := FALSE;
   END_IF;
END_REGION

REGION Network 15: Falha retorno valvulas
   #TON_FalhaRetornoValvProd1(IN := #AcionaValvProd1 AND NOT #RetValvProd1, PT := T#5s);   // TON
   IF #TON_FalhaRetornoValvProd1.Q THEN #FalhaValvProd1 := TRUE; END_IF;
   #TON_FalhaRetornoValvProd2(IN := #AcionaValvProd2 AND NOT #RetValvProd2, PT := T#5s);   // TON
   IF #TON_FalhaRetornoValvProd2.Q THEN #FalhaValvProd2 := TRUE; END_IF;
   IF "ResetGeral" THEN
       #FalhaValvProd1 := FALSE;
       #FalhaValvProd2 := FALSE;
   END_IF;
END_REGION

REGION Network 16: Status Bomba (0 - Sem alarmes; 1 - Bomba ligada; 2 - Bomba em alarme; 3 - Bomba em manutenção)
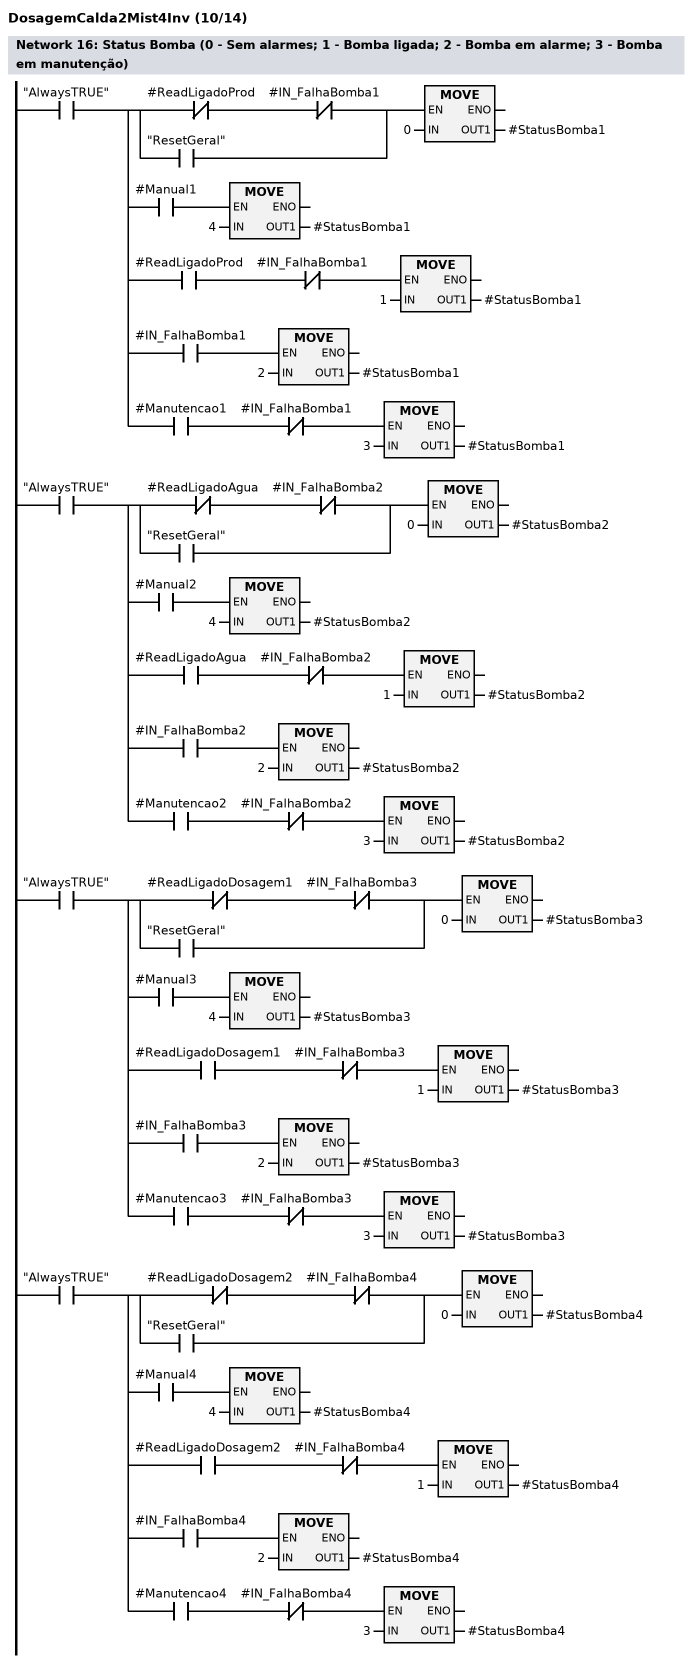
   RUNG wire#powerrail
      Contact( "AlwaysTRUE" )
      wire#w1
      I_Contact( #ReadLigadoProd )
      I_Contact( #IN_FalhaBomba1 )
      wire#w2
      Move(in := 0, out1 => #StatusBomba1)
   END_RUNG
   RUNG wire#w1
      Contact( "ResetGeral" )
   END_RUNG wire#w2
   RUNG wire#w1
      Contact( #Manual1 )
      Move(in := 4, out1 => #StatusBomba1)
   END_RUNG
   RUNG wire#w1
      Contact( #ReadLigadoProd )
      I_Contact( #IN_FalhaBomba1 )
      Move(in := 1, out1 => #StatusBomba1)
   END_RUNG
   RUNG wire#w1
      Contact( #IN_FalhaBomba1 )
      Move(in := 2, out1 => #StatusBomba1)
   END_RUNG
   RUNG wire#w1
      Contact( #Manutencao1 )
      I_Contact( #IN_FalhaBomba1 )
      Move(in := 3, out1 => #StatusBomba1)
   END_RUNG
   RUNG wire#powerrail
      Contact( "AlwaysTRUE" )
      wire#w3
      I_Contact( #ReadLigadoAgua )
      I_Contact( #IN_FalhaBomba2 )
      wire#w4
      Move(in := 0, out1 => #StatusBomba2)
   END_RUNG
   RUNG wire#w3
      Contact( "ResetGeral" )
   END_RUNG wire#w4
   RUNG wire#w3
      Contact( #Manual2 )
      Move(in := 4, out1 => #StatusBomba2)
   END_RUNG
   RUNG wire#w3
      Contact( #ReadLigadoAgua )
      I_Contact( #IN_FalhaBomba2 )
      Move(in := 1, out1 => #StatusBomba2)
   END_RUNG
   RUNG wire#w3
      Contact( #IN_FalhaBomba2 )
      Move(in := 2, out1 => #StatusBomba2)
   END_RUNG
   RUNG wire#w3
      Contact( #Manutencao2 )
      I_Contact( #IN_FalhaBomba2 )
      Move(in := 3, out1 => #StatusBomba2)
   END_RUNG
   RUNG wire#powerrail
      Contact( "AlwaysTRUE" )
      wire#w5
      I_Contact( #ReadLigadoDosagem1 )
      I_Contact( #IN_FalhaBomba3 )
      wire#w6
      Move(in := 0, out1 => #StatusBomba3)
   END_RUNG
   RUNG wire#w5
      Contact( "ResetGeral" )
   END_RUNG wire#w6
   RUNG wire#w5
      Contact( #Manual3 )
      Move(in := 4, out1 => #StatusBomba3)
   END_RUNG
   RUNG wire#w5
      Contact( #ReadLigadoDosagem1 )
      I_Contact( #IN_FalhaBomba3 )
      Move(in := 1, out1 => #StatusBomba3)
   END_RUNG
   RUNG wire#w5
      Contact( #IN_FalhaBomba3 )
      Move(in := 2, out1 => #StatusBomba3)
   END_RUNG
   RUNG wire#w5
      Contact( #Manutencao3 )
      I_Contact( #IN_FalhaBomba3 )
      Move(in := 3, out1 => #StatusBomba3)
   END_RUNG
   RUNG wire#powerrail
      Contact( "AlwaysTRUE" )
      wire#w7
      I_Contact( #ReadLigadoDosagem2 )
      I_Contact( #IN_FalhaBomba4 )
      wire#w8
      Move(in := 0, out1 => #StatusBomba4)
   END_RUNG
   RUNG wire#w7
      Contact( "ResetGeral" )
   END_RUNG wire#w8
   RUNG wire#w7
      Contact( #Manual4 )
      Move(in := 4, out1 => #StatusBomba4)
   END_RUNG
   RUNG wire#w7
      Contact( #ReadLigadoDosagem2 )
      I_Contact( #IN_FalhaBomba4 )
      Move(in := 1, out1 => #StatusBomba4)
   END_RUNG
   RUNG wire#w7
      Contact( #IN_FalhaBomba4 )
      Move(in := 2, out1 => #StatusBomba4)
   END_RUNG
   RUNG wire#w7
      Contact( #Manutencao4 )
      I_Contact( #IN_FalhaBomba4 )
      Move(in := 3, out1 => #StatusBomba4)
   END_RUNG
   // the same network as SCL:
   IF "AlwaysTRUE" AND ((NOT #ReadLigadoProd AND NOT #IN_FalhaBomba1) OR "ResetGeral") THEN
       #StatusBomba1 := 0;
   END_IF;
   IF "AlwaysTRUE" AND #Manual1 THEN #StatusBomba1 := 4; END_IF;
   IF "AlwaysTRUE" AND #ReadLigadoProd AND NOT #IN_FalhaBomba1 THEN #StatusBomba1 := 1; END_IF;
   IF "AlwaysTRUE" AND #IN_FalhaBomba1 THEN #StatusBomba1 := 2; END_IF;
   IF "AlwaysTRUE" AND #Manutencao1 AND NOT #IN_FalhaBomba1 THEN #StatusBomba1 := 3; END_IF;
   IF "AlwaysTRUE" AND ((NOT #ReadLigadoAgua AND NOT #IN_FalhaBomba2) OR "ResetGeral") THEN
       #StatusBomba2 := 0;
   END_IF;
   IF "AlwaysTRUE" AND #Manual2 THEN #StatusBomba2 := 4; END_IF;
   IF "AlwaysTRUE" AND #ReadLigadoAgua AND NOT #IN_FalhaBomba2 THEN #StatusBomba2 := 1; END_IF;
   IF "AlwaysTRUE" AND #IN_FalhaBomba2 THEN #StatusBomba2 := 2; END_IF;
   IF "AlwaysTRUE" AND #Manutencao2 AND NOT #IN_FalhaBomba2 THEN #StatusBomba2 := 3; END_IF;
   IF "AlwaysTRUE" AND ((NOT #ReadLigadoDosagem1 AND NOT #IN_FalhaBomba3) OR "ResetGeral") THEN
       #StatusBomba3 := 0;
   END_IF;
   IF "AlwaysTRUE" AND #Manual3 THEN #StatusBomba3 := 4; END_IF;
   IF "AlwaysTRUE" AND #ReadLigadoDosagem1 AND NOT #IN_FalhaBomba3 THEN #StatusBomba3 := 1; END_IF;
   IF "AlwaysTRUE" AND #IN_FalhaBomba3 THEN #StatusBomba3 := 2; END_IF;
   IF "AlwaysTRUE" AND #Manutencao3 AND NOT #IN_FalhaBomba3 THEN #StatusBomba3 := 3; END_IF;
   IF "AlwaysTRUE" AND ((NOT #ReadLigadoDosagem2 AND NOT #IN_FalhaBomba4) OR "ResetGeral") THEN
       #StatusBomba4 := 0;
   END_IF;
   IF "AlwaysTRUE" AND #Manual4 THEN #StatusBomba4 := 4; END_IF;
   IF "AlwaysTRUE" AND #ReadLigadoDosagem2 AND NOT #IN_FalhaBomba4 THEN #StatusBomba4 := 1; END_IF;
   IF "AlwaysTRUE" AND #IN_FalhaBomba4 THEN #StatusBomba4 := 2; END_IF;
   IF "AlwaysTRUE" AND #Manutencao4 AND NOT #IN_FalhaBomba4 THEN #StatusBomba4 := 3; END_IF;
END_REGION

REGION Network 17: Icone Bomba (0 - Automatico; 1 - Manual; 2 - Manutenção)
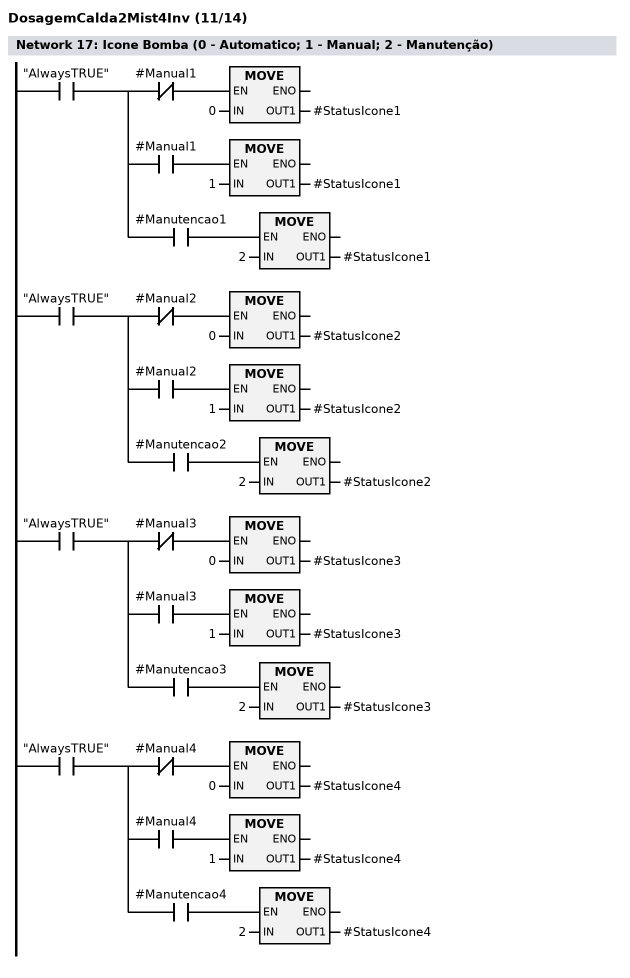
   RUNG wire#powerrail
      Contact( "AlwaysTRUE" )
      wire#w1
      I_Contact( #Manual1 )
      Move(in := 0, out1 => #StatusIcone1)
   END_RUNG
   RUNG wire#w1
      Contact( #Manual1 )
      Move(in := 1, out1 => #StatusIcone1)
   END_RUNG
   RUNG wire#w1
      Contact( #Manutencao1 )
      Move(in := 2, out1 => #StatusIcone1)
   END_RUNG
   RUNG wire#powerrail
      Contact( "AlwaysTRUE" )
      wire#w2
      I_Contact( #Manual2 )
      Move(in := 0, out1 => #StatusIcone2)
   END_RUNG
   RUNG wire#w2
      Contact( #Manual2 )
      Move(in := 1, out1 => #StatusIcone2)
   END_RUNG
   RUNG wire#w2
      Contact( #Manutencao2 )
      Move(in := 2, out1 => #StatusIcone2)
   END_RUNG
   RUNG wire#powerrail
      Contact( "AlwaysTRUE" )
      wire#w3
      I_Contact( #Manual3 )
      Move(in := 0, out1 => #StatusIcone3)
   END_RUNG
   RUNG wire#w3
      Contact( #Manual3 )
      Move(in := 1, out1 => #StatusIcone3)
   END_RUNG
   RUNG wire#w3
      Contact( #Manutencao3 )
      Move(in := 2, out1 => #StatusIcone3)
   END_RUNG
   RUNG wire#powerrail
      Contact( "AlwaysTRUE" )
      wire#w4
      I_Contact( #Manual4 )
      Move(in := 0, out1 => #StatusIcone4)
   END_RUNG
   RUNG wire#w4
      Contact( #Manual4 )
      Move(in := 1, out1 => #StatusIcone4)
   END_RUNG
   RUNG wire#w4
      Contact( #Manutencao4 )
      Move(in := 2, out1 => #StatusIcone4)
   END_RUNG
   // the same network as SCL:
   IF "AlwaysTRUE" AND NOT #Manual1 THEN #StatusIcone1 := 0; END_IF;
   IF "AlwaysTRUE" AND #Manual1 THEN #StatusIcone1 := 1; END_IF;
   IF "AlwaysTRUE" AND #Manutencao1 THEN #StatusIcone1 := 2; END_IF;
   IF "AlwaysTRUE" AND NOT #Manual2 THEN #StatusIcone2 := 0; END_IF;
   IF "AlwaysTRUE" AND #Manual2 THEN #StatusIcone2 := 1; END_IF;
   IF "AlwaysTRUE" AND #Manutencao2 THEN #StatusIcone2 := 2; END_IF;
   IF "AlwaysTRUE" AND NOT #Manual3 THEN #StatusIcone3 := 0; END_IF;
   IF "AlwaysTRUE" AND #Manual3 THEN #StatusIcone3 := 1; END_IF;
   IF "AlwaysTRUE" AND #Manutencao3 THEN #StatusIcone3 := 2; END_IF;
   IF "AlwaysTRUE" AND NOT #Manual4 THEN #StatusIcone4 := 0; END_IF;
   IF "AlwaysTRUE" AND #Manual4 THEN #StatusIcone4 := 1; END_IF;
   IF "AlwaysTRUE" AND #Manutencao4 THEN #StatusIcone4 := 2; END_IF;
END_REGION

REGION Network 18: Somatoria para diario e totalizadores 1
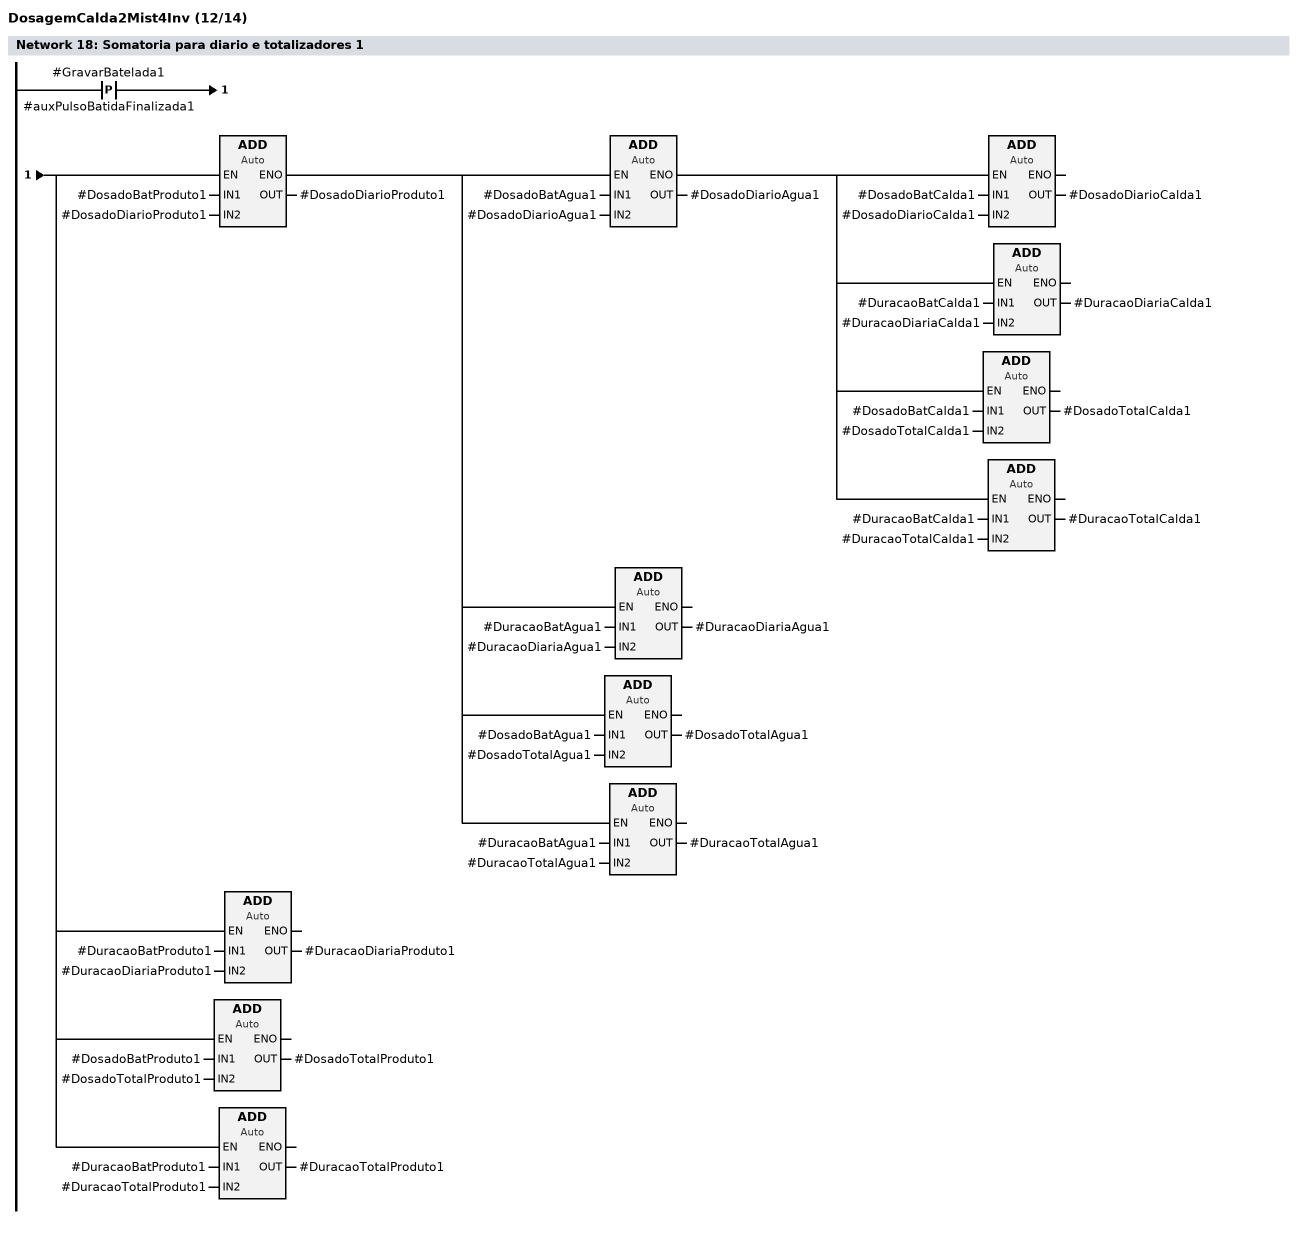
   RUNG wire#powerrail
      P_Contact(operand := #GravarBatelada1, bit := #auxPulsoBatidaFinalizada1)
      wire#w1
      Add(in1 := #DosadoBatProduto1, in2 := #DosadoDiarioProduto1, out => #DosadoDiarioProduto1)
      wire#w2
      Add(in1 := #DosadoBatAgua1, in2 := #DosadoDiarioAgua1, out => #DosadoDiarioAgua1)
      wire#w3
      Add(in1 := #DosadoBatCalda1, in2 := #DosadoDiarioCalda1, out => #DosadoDiarioCalda1)
   END_RUNG
   RUNG wire#w3
      Add(in1 := #DuracaoBatCalda1, in2 := #DuracaoDiariaCalda1, out => #DuracaoDiariaCalda1)
   END_RUNG
   RUNG wire#w3
      Add(in1 := #DosadoBatCalda1, in2 := #DosadoTotalCalda1, out => #DosadoTotalCalda1)
   END_RUNG
   RUNG wire#w3
      Add(in1 := #DuracaoBatCalda1, in2 := #DuracaoTotalCalda1, out => #DuracaoTotalCalda1)
   END_RUNG
   RUNG wire#w2
      Add(in1 := #DuracaoBatAgua1, in2 := #DuracaoDiariaAgua1, out => #DuracaoDiariaAgua1)
   END_RUNG
   RUNG wire#w2
      Add(in1 := #DosadoBatAgua1, in2 := #DosadoTotalAgua1, out => #DosadoTotalAgua1)
   END_RUNG
   RUNG wire#w2
      Add(in1 := #DuracaoBatAgua1, in2 := #DuracaoTotalAgua1, out => #DuracaoTotalAgua1)
   END_RUNG
   RUNG wire#w1
      Add(in1 := #DuracaoBatProduto1, in2 := #DuracaoDiariaProduto1, out => #DuracaoDiariaProduto1)
   END_RUNG
   RUNG wire#w1
      Add(in1 := #DosadoBatProduto1, in2 := #DosadoTotalProduto1, out => #DosadoTotalProduto1)
   END_RUNG
   RUNG wire#w1
      Add(in1 := #DuracaoBatProduto1, in2 := #DuracaoTotalProduto1, out => #DuracaoTotalProduto1)
   END_RUNG
   // the same network as SCL:
   #_w1 := #GravarBatelada1 AND NOT #auxPulsoBatidaFinalizada1;   // rising edge of #GravarBatelada1
   #auxPulsoBatidaFinalizada1 := #GravarBatelada1;
   IF #_w1 THEN
       #DosadoDiarioProduto1 := #DosadoBatProduto1 + #DosadoDiarioProduto1;
       #DosadoDiarioAgua1 := #DosadoBatAgua1 + #DosadoDiarioAgua1;
       #DosadoDiarioCalda1 := #DosadoBatCalda1 + #DosadoDiarioCalda1;
       #DuracaoDiariaCalda1 := #DuracaoBatCalda1 + #DuracaoDiariaCalda1;
       #DosadoTotalCalda1 := #DosadoBatCalda1 + #DosadoTotalCalda1;
       #DuracaoTotalCalda1 := #DuracaoBatCalda1 + #DuracaoTotalCalda1;
       #DuracaoDiariaAgua1 := #DuracaoBatAgua1 + #DuracaoDiariaAgua1;
       #DosadoTotalAgua1 := #DosadoBatAgua1 + #DosadoTotalAgua1;
       #DuracaoTotalAgua1 := #DuracaoBatAgua1 + #DuracaoTotalAgua1;
       #DuracaoDiariaProduto1 := #DuracaoBatProduto1 + #DuracaoDiariaProduto1;
       #DosadoTotalProduto1 := #DosadoBatProduto1 + #DosadoTotalProduto1;
       #DuracaoTotalProduto1 := #DuracaoBatProduto1 + #DuracaoTotalProduto1;
   END_IF;
END_REGION

REGION Network 19: Somatoria para diario e totalizadores 2
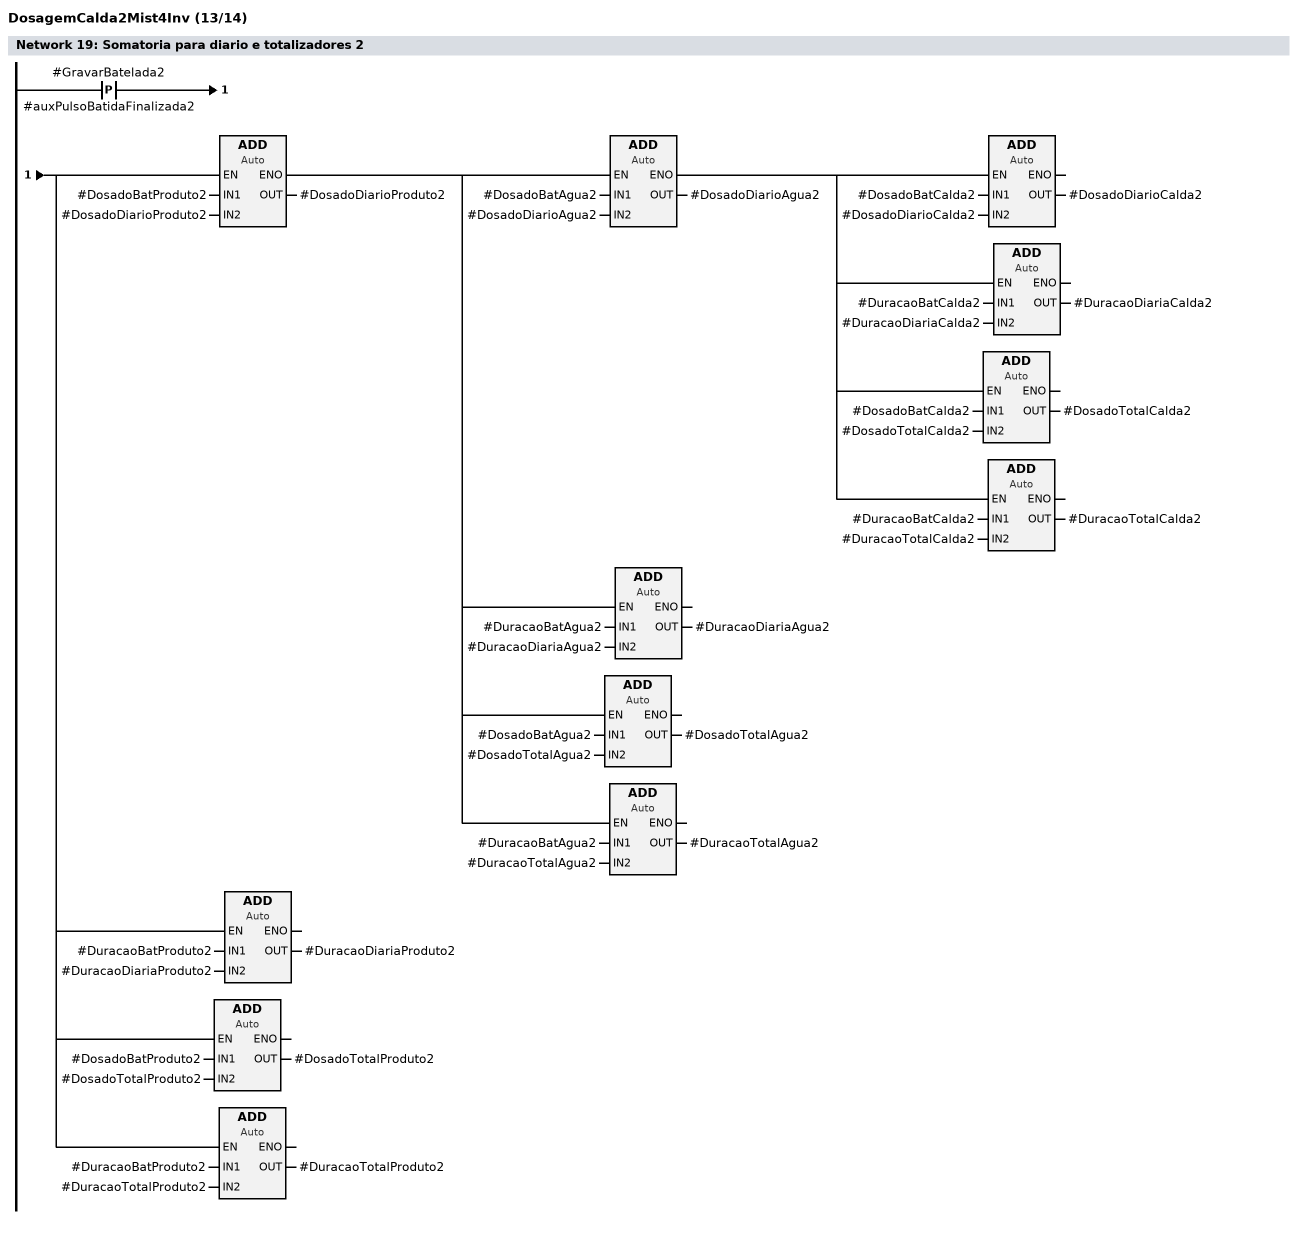
   RUNG wire#powerrail
      P_Contact(operand := #GravarBatelada2, bit := #auxPulsoBatidaFinalizada2)
      wire#w1
      Add(in1 := #DosadoBatProduto2, in2 := #DosadoDiarioProduto2, out => #DosadoDiarioProduto2)
      wire#w2
      Add(in1 := #DosadoBatAgua2, in2 := #DosadoDiarioAgua2, out => #DosadoDiarioAgua2)
      wire#w3
      Add(in1 := #DosadoBatCalda2, in2 := #DosadoDiarioCalda2, out => #DosadoDiarioCalda2)
   END_RUNG
   RUNG wire#w3
      Add(in1 := #DuracaoBatCalda2, in2 := #DuracaoDiariaCalda2, out => #DuracaoDiariaCalda2)
   END_RUNG
   RUNG wire#w3
      Add(in1 := #DosadoBatCalda2, in2 := #DosadoTotalCalda2, out => #DosadoTotalCalda2)
   END_RUNG
   RUNG wire#w3
      Add(in1 := #DuracaoBatCalda2, in2 := #DuracaoTotalCalda2, out => #DuracaoTotalCalda2)
   END_RUNG
   RUNG wire#w2
      Add(in1 := #DuracaoBatAgua2, in2 := #DuracaoDiariaAgua2, out => #DuracaoDiariaAgua2)
   END_RUNG
   RUNG wire#w2
      Add(in1 := #DosadoBatAgua2, in2 := #DosadoTotalAgua2, out => #DosadoTotalAgua2)
   END_RUNG
   RUNG wire#w2
      Add(in1 := #DuracaoBatAgua2, in2 := #DuracaoTotalAgua2, out => #DuracaoTotalAgua2)
   END_RUNG
   RUNG wire#w1
      Add(in1 := #DuracaoBatProduto2, in2 := #DuracaoDiariaProduto2, out => #DuracaoDiariaProduto2)
   END_RUNG
   RUNG wire#w1
      Add(in1 := #DosadoBatProduto2, in2 := #DosadoTotalProduto2, out => #DosadoTotalProduto2)
   END_RUNG
   RUNG wire#w1
      Add(in1 := #DuracaoBatProduto2, in2 := #DuracaoTotalProduto2, out => #DuracaoTotalProduto2)
   END_RUNG
   // the same network as SCL:
   #_w1 := #GravarBatelada2 AND NOT #auxPulsoBatidaFinalizada2;   // rising edge of #GravarBatelada2
   #auxPulsoBatidaFinalizada2 := #GravarBatelada2;
   IF #_w1 THEN
       #DosadoDiarioProduto2 := #DosadoBatProduto2 + #DosadoDiarioProduto2;
       #DosadoDiarioAgua2 := #DosadoBatAgua2 + #DosadoDiarioAgua2;
       #DosadoDiarioCalda2 := #DosadoBatCalda2 + #DosadoDiarioCalda2;
       #DuracaoDiariaCalda2 := #DuracaoBatCalda2 + #DuracaoDiariaCalda2;
       #DosadoTotalCalda2 := #DosadoBatCalda2 + #DosadoTotalCalda2;
       #DuracaoTotalCalda2 := #DuracaoBatCalda2 + #DuracaoTotalCalda2;
       #DuracaoDiariaAgua2 := #DuracaoBatAgua2 + #DuracaoDiariaAgua2;
       #DosadoTotalAgua2 := #DosadoBatAgua2 + #DosadoTotalAgua2;
       #DuracaoTotalAgua2 := #DuracaoBatAgua2 + #DuracaoTotalAgua2;
       #DuracaoDiariaProduto2 := #DuracaoBatProduto2 + #DuracaoDiariaProduto2;
       #DosadoTotalProduto2 := #DosadoBatProduto2 + #DosadoTotalProduto2;
       #DuracaoTotalProduto2 := #DuracaoBatProduto2 + #DuracaoTotalProduto2;
   END_IF;
END_REGION

REGION Network 20: Trigger / reset para relatorio diario e totalizador
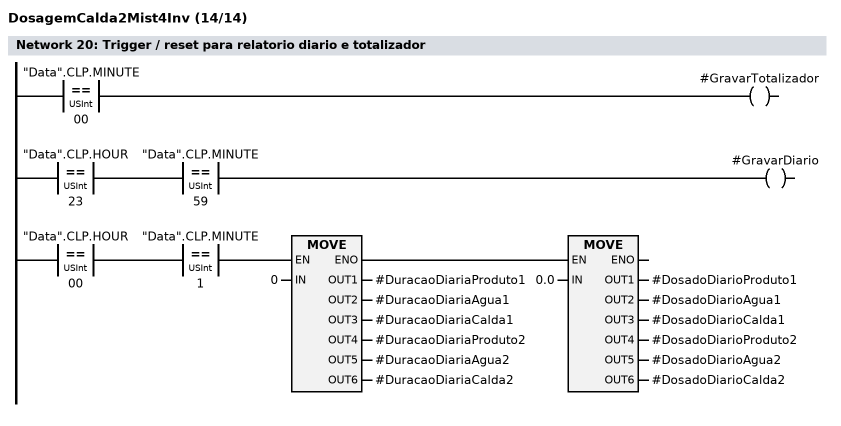
   RUNG wire#powerrail
      { S7_Templates := "SrcType := USInt" } EQ_Contact(in1 := "Data".CLP.MINUTE, in2 := 00)
      Coil( #GravarTotalizador )
   END_RUNG
   RUNG wire#powerrail
      { S7_Templates := "SrcType := USInt" } EQ_Contact(in1 := "Data".CLP.HOUR, in2 := 23)
      { S7_Templates := "SrcType := USInt" } EQ_Contact(in1 := "Data".CLP.MINUTE, in2 := 59)
      Coil( #GravarDiario )
   END_RUNG
   RUNG wire#powerrail
      { S7_Templates := "SrcType := USInt" } EQ_Contact(in1 := "Data".CLP.HOUR, in2 := 00)
      { S7_Templates := "SrcType := USInt" } EQ_Contact(in1 := "Data".CLP.MINUTE, in2 := 1)
      Move(in := 0, out1 => #DuracaoDiariaProduto1, out2 => #DuracaoDiariaAgua1, out3 => #DuracaoDiariaCalda1, out4 => #DuracaoDiariaProduto2, out5 => #DuracaoDiariaAgua2, out6 => #DuracaoDiariaCalda2)
      Move(in := 0.0, out1 => #DosadoDiarioProduto1, out2 => #DosadoDiarioAgua1, out3 => #DosadoDiarioCalda1, out4 => #DosadoDiarioProduto2, out5 => #DosadoDiarioAgua2, out6 => #DosadoDiarioCalda2)
   END_RUNG
   // the same network as SCL:
   #GravarTotalizador := "Data".CLP.MINUTE = 00;
   #GravarDiario := ("Data".CLP.HOUR = 23) AND ("Data".CLP.MINUTE = 59);
   IF ("Data".CLP.HOUR = 00) AND ("Data".CLP.MINUTE = 1) THEN
       #DuracaoDiariaProduto1 := 0;
       #DuracaoDiariaAgua1 := 0;
       #DuracaoDiariaCalda1 := 0;
       #DuracaoDiariaProduto2 := 0;
       #DuracaoDiariaAgua2 := 0;
       #DuracaoDiariaCalda2 := 0;
       #DosadoDiarioProduto1 := 0.0;
       #DosadoDiarioAgua1 := 0.0;
       #DosadoDiarioCalda1 := 0.0;
       #DosadoDiarioProduto2 := 0.0;
       #DosadoDiarioAgua2 := 0.0;
       #DosadoDiarioCalda2 := 0.0;
   END_IF;
END_REGION
END_FUNCTION_BLOCK

FUNCTION_BLOCK "DosagemMisturador"   // FB101, LAD
{ S7_Optimized_Access := 'TRUE' }
VERSION : 0.1
   VAR_INPUT
      SistemaHabilitado : Bool;
      Emergencia : Bool;
      SinalDosagem : Bool;
      PulsoMedidor : Bool;
      VolumePulso_ml : Real := 1.0;
      RetValvulaAberta : Bool;
      SP_Quant : Real;
      SP_AjusteFino : Real;
      SP_Corte : Real;
      SP_TempoMax : Time;
      SP_TempMistSeca : Time;
      SP_FreqMax : Real;
      SP_FreqMin : Real;
      IN_FalhaBomba : Bool;
      IN_InversorError : Bool;
      ReadLigado : Bool;
   END_VAR
   VAR_OUTPUT
      LigaBomba : Bool;
      LigarValvula : Bool;
      FreqAtual : Real;
      FalhaBomba : Bool;
      FalhaValvula : Bool;
      FalhaTempoMax : Bool;
   END_VAR
   VAR_IN_OUT
      DosadoDiario : Real;
      DuracaoDiaria : Real;
      DosadoTotal : LReal;
      DuracaoTotal : LReal;
   END_VAR
   VAR RETAIN
      TON_EstabilizaBalanca : TON_TIME;
      QuantAlvo : Real;
      auxPulsoSinalDosagem : Bool;
      TON_MisturaSeca : TON_TIME;
      auxSetSinalDosagem : Bool;
      HabilitadoDosagem : Bool;
      TON_AbreContatora : TON_TIME;
      QuantAjuste : Real;
      auxPulsoClock1HZ : Bool;
      auxPulsoBatidaFinalizada : Bool;
      auxPulsoMedVazao : Bool;
      QuantDosadaAux : Real;
      auxPulsoLigarBomba : Bool;
      AlvoAjusteFino : Real;
      AlvoDosagem : Real;
      TON_FalhaRetornoBomba : TON_TIME;
      TON_FalhaValvula : TON_TIME;
      TON_ResetSinalFabrica : TON_TIME;
      auxTempoMax : DInt;
      TOF_MantemRegistro : TOF_TIME;
      TON_FaltaFluxo : TON_TIME;
      auxTempoMistSeca : DInt;
      auxTempoMisturaSecaDecorrido : DInt;
      TempoMaxRestante : DInt;
      TON_RetardoGravaBatida : TON_TIME;
      auxGravaBatida : Bool;
      DuracaoBat : Real;
      DosadoBat : Real;
      StatusBomba : Int;
      StatusIcone : Int;
      BatidaFinalizada : Bool;
      GravarBatida : Bool;
      auxNegaReadLigado : Bool;
      Manual : Bool;
      LigaManual : Bool;
      Manutencao : Bool;
      TOF_DelayGravarBatida : TOF_TIME;
      TempoMistSecaRestante : DInt;
      TON_DelaySalvaBat : TON_TIME;
      VolumePulso_l : Real;
      AcumuladoIntegracao : Real;
      nReadLigado : Bool;
   END_VAR
   VAR_TEMP   // added for the SCL form of the ladder/FBD networks
      _w1 : Bool;
      _w2 : Bool;
      _w3 : Bool;
   END_VAR
BEGIN

REGION Network 1: Tempo de mistura seca / tempo maximo
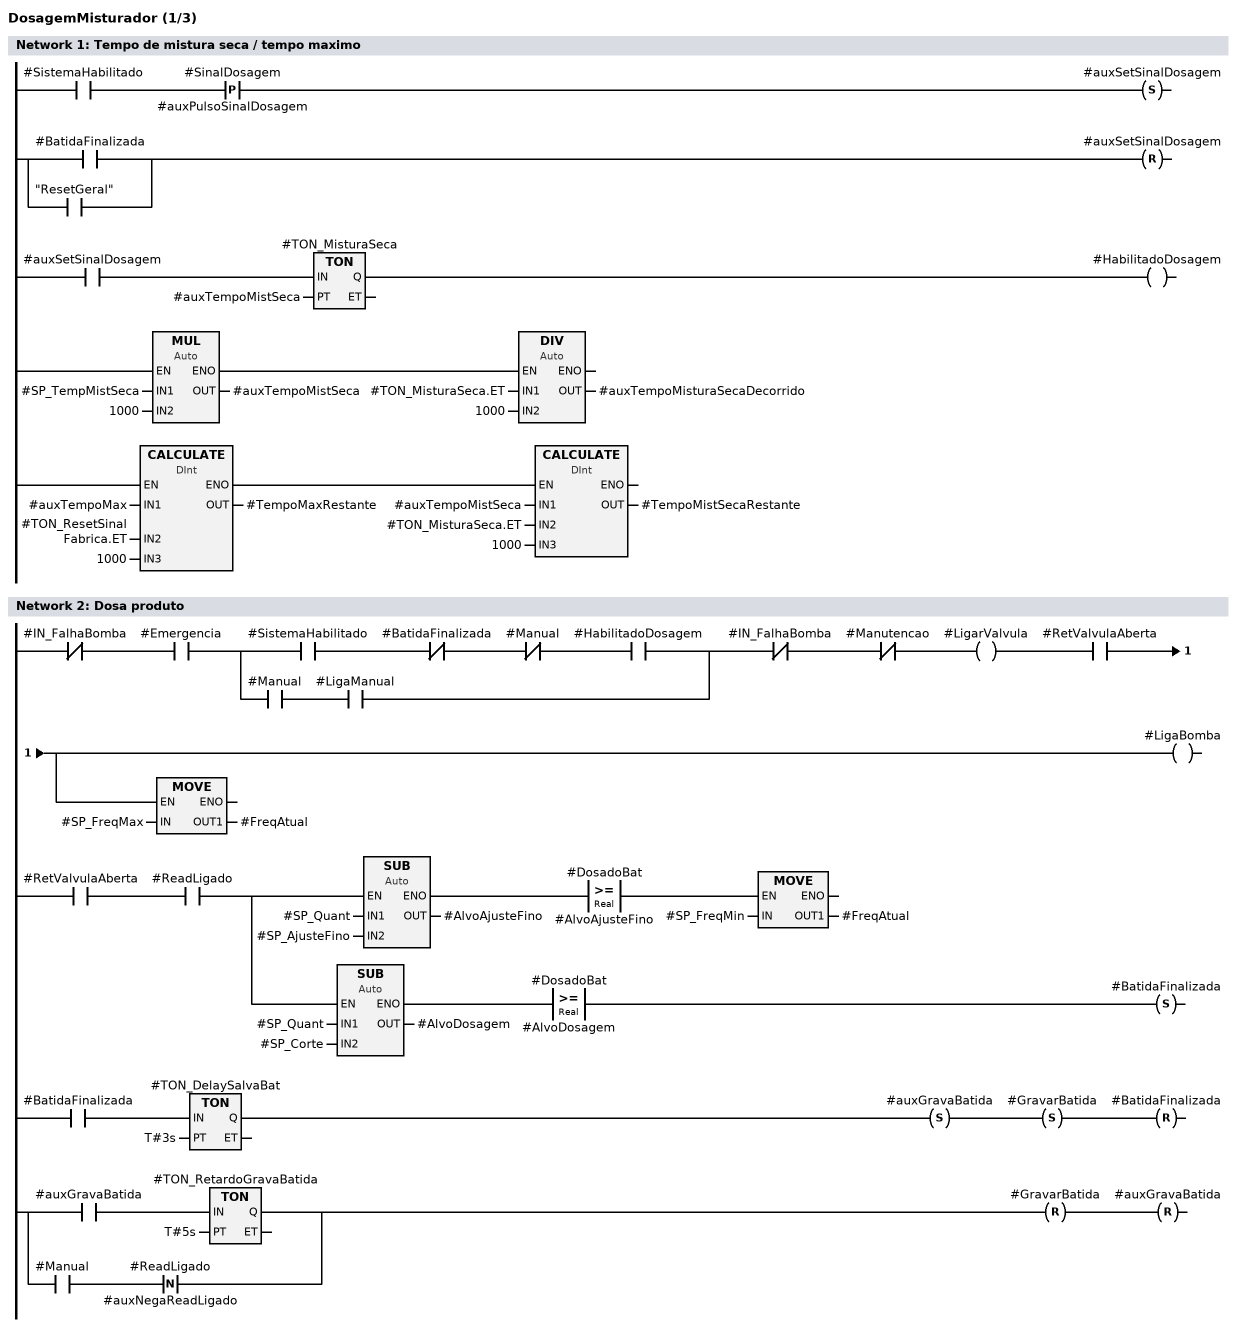
   #_w1 := #SistemaHabilitado AND #SinalDosagem AND NOT #auxPulsoSinalDosagem;   // rising edge of #SinalDosagem
   #auxPulsoSinalDosagem := #SinalDosagem;
   IF #_w1 THEN #auxSetSinalDosagem := TRUE; END_IF;
   IF #BatidaFinalizada OR "ResetGeral" THEN #auxSetSinalDosagem := FALSE; END_IF;
   #TON_MisturaSeca(IN := #auxSetSinalDosagem, PT := #auxTempoMistSeca);   // TON
   #HabilitadoDosagem := #TON_MisturaSeca.Q;
   #auxTempoMistSeca := #SP_TempMistSeca * 1000;
   #auxTempoMisturaSecaDecorrido := #TON_MisturaSeca.ET / 1000;
   #TempoMaxRestante := ((#auxTempoMax - #TON_ResetSinalFabrica.ET) / 1000);
   #TempoMistSecaRestante := ((#auxTempoMistSeca - #TON_MisturaSeca.ET) / 1000);
END_REGION

REGION Network 2: Dosa produto
   #LigarValvula := NOT #IN_FalhaBomba AND #Emergencia AND ((#SistemaHabilitado AND NOT #BatidaFinalizada AND NOT #Manual AND #HabilitadoDosagem) OR (#Manual AND #LigaManual)) AND NOT #IN_FalhaBomba AND NOT #Manutencao;
   #LigaBomba := #LigarValvula AND #RetValvulaAberta;
   IF #LigaBomba THEN #FreqAtual := #SP_FreqMax; END_IF;
   #_w1 := #RetValvulaAberta AND #ReadLigado;
   IF #_w1 THEN #AlvoAjusteFino := #SP_Quant - #SP_AjusteFino; END_IF;
   IF #_w1 AND (#DosadoBat >= #AlvoAjusteFino) THEN #FreqAtual := #SP_FreqMin; END_IF;
   IF #_w1 THEN #AlvoDosagem := #SP_Quant - #SP_Corte; END_IF;
   IF #_w1 AND (#DosadoBat >= #AlvoDosagem) THEN #BatidaFinalizada := TRUE; END_IF;
   #TON_DelaySalvaBat(IN := #BatidaFinalizada, PT := T#3s);   // TON
   IF #TON_DelaySalvaBat.Q THEN
       #auxGravaBatida := TRUE;
       #GravarBatida := TRUE;
       #BatidaFinalizada := FALSE;
   END_IF;
   #TON_RetardoGravaBatida(IN := #auxGravaBatida, PT := T#5s);   // TON
   #_w2 := #Manual AND NOT #ReadLigado AND #auxNegaReadLigado;   // falling edge of #ReadLigado
   #auxNegaReadLigado := #ReadLigado;
   IF #TON_RetardoGravaBatida.Q OR #_w2 THEN
       #GravarBatida := FALSE;
       #auxGravaBatida := FALSE;
   END_IF;
END_REGION

REGION Network 3: Registra Acumulados
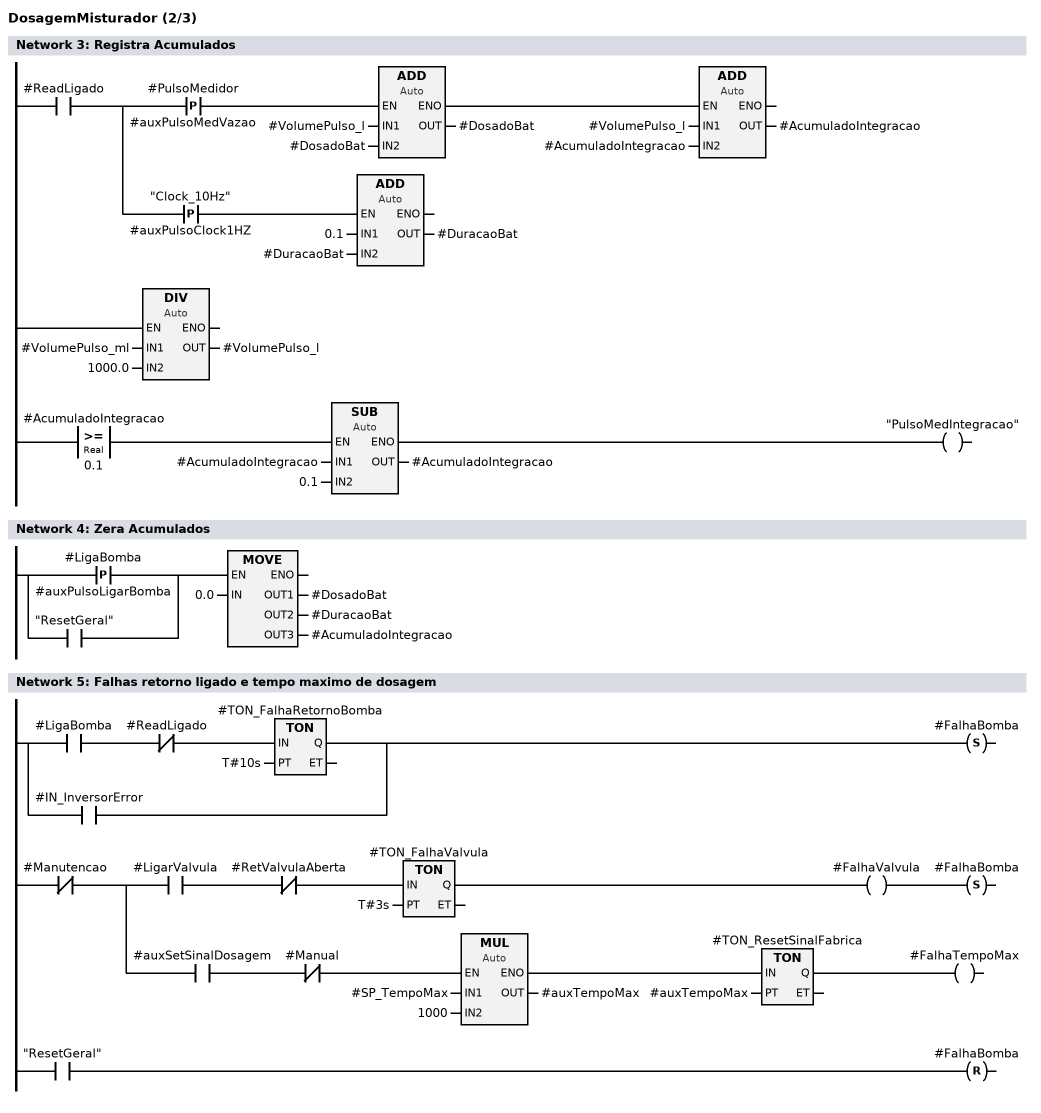
   RUNG wire#powerrail
      Contact( #ReadLigado )
      wire#w1
      P_Contact(operand := #PulsoMedidor, bit := #auxPulsoMedVazao)
      Add(in1 := #VolumePulso_l, in2 := #DosadoBat, out => #DosadoBat)
      Add(in1 := #VolumePulso_l, in2 := #AcumuladoIntegracao, out => #AcumuladoIntegracao)
   END_RUNG
   RUNG wire#w1
      P_Contact(operand := "Clock_10Hz", bit := #auxPulsoClock1HZ)
      Add(in1 := 0.1, in2 := #DuracaoBat, out => #DuracaoBat)
   END_RUNG
   RUNG wire#powerrail
      Div(in1 := #VolumePulso_ml, in2 := 1000.0, out => #VolumePulso_l)
   END_RUNG
   RUNG wire#powerrail
      { S7_Templates := "SrcType := Real" } GE_Contact(in1 := #AcumuladoIntegracao, in2 := 0.1)
      Sub(in1 := #AcumuladoIntegracao, in2 := 0.1, out => #AcumuladoIntegracao)
      Coil( "PulsoMedIntegracao" )
   END_RUNG
   // the same network as SCL:
   #_w1 := #ReadLigado AND #PulsoMedidor AND NOT #auxPulsoMedVazao;   // rising edge of #PulsoMedidor
   #auxPulsoMedVazao := #PulsoMedidor;
   IF #_w1 THEN
       #DosadoBat := #VolumePulso_l + #DosadoBat;
       #AcumuladoIntegracao := #VolumePulso_l + #AcumuladoIntegracao;
   END_IF;
   #_w2 := #ReadLigado AND "Clock_10Hz" AND NOT #auxPulsoClock1HZ;   // rising edge of "Clock_10Hz"
   #auxPulsoClock1HZ := "Clock_10Hz";
   IF #_w2 THEN #DuracaoBat := 0.1 + #DuracaoBat; END_IF;
   #VolumePulso_l := #VolumePulso_ml / 1000.0;
   #_w3 := #AcumuladoIntegracao >= 0.1;
   IF #_w3 THEN #AcumuladoIntegracao := #AcumuladoIntegracao - 0.1; END_IF;
   "PulsoMedIntegracao" := #_w3;
END_REGION

REGION Network 4: Zera Acumulados
   RUNG wire#powerrail
      P_Contact(operand := #LigaBomba, bit := #auxPulsoLigarBomba)
      wire#w1
      Move(in := 0.0, out1 => #DosadoBat, out2 => #DuracaoBat, out3 => #AcumuladoIntegracao)
   END_RUNG
   RUNG wire#powerrail
      Contact( "ResetGeral" )
   END_RUNG wire#w1
   // the same network as SCL:
   #_w1 := #LigaBomba AND NOT #auxPulsoLigarBomba;   // rising edge of #LigaBomba
   #auxPulsoLigarBomba := #LigaBomba;
   IF #_w1 OR "ResetGeral" THEN
       #DosadoBat := 0.0;
       #DuracaoBat := 0.0;
       #AcumuladoIntegracao := 0.0;
   END_IF;
END_REGION

REGION Network 5: Falhas retorno ligado e tempo maximo de dosagem
   #TON_FalhaRetornoBomba(IN := #LigaBomba AND NOT #ReadLigado, PT := T#10s);   // TON
   IF #TON_FalhaRetornoBomba.Q OR #IN_InversorError THEN #FalhaBomba := TRUE; END_IF;
   #TON_FalhaValvula(IN := NOT #Manutencao AND #LigarValvula AND NOT #RetValvulaAberta, PT := T#3s);   // TON
   #FalhaValvula := #TON_FalhaValvula.Q;
   IF #TON_FalhaValvula.Q THEN #FalhaBomba := TRUE; END_IF;
   #_w1 := NOT #Manutencao AND #auxSetSinalDosagem AND NOT #Manual;
   IF #_w1 THEN #auxTempoMax := #SP_TempoMax * 1000; END_IF;
   #TON_ResetSinalFabrica(IN := #_w1, PT := #auxTempoMax);   // TON
   #FalhaTempoMax := #TON_ResetSinalFabrica.Q;
   IF "ResetGeral" THEN #FalhaBomba := FALSE; END_IF;
END_REGION

REGION Network 6: Status Bomba (0 - Sem alarmes; 1 - Bomba ligada; 2 - Bomba em alarme; 3 - Bomba em manutenção)
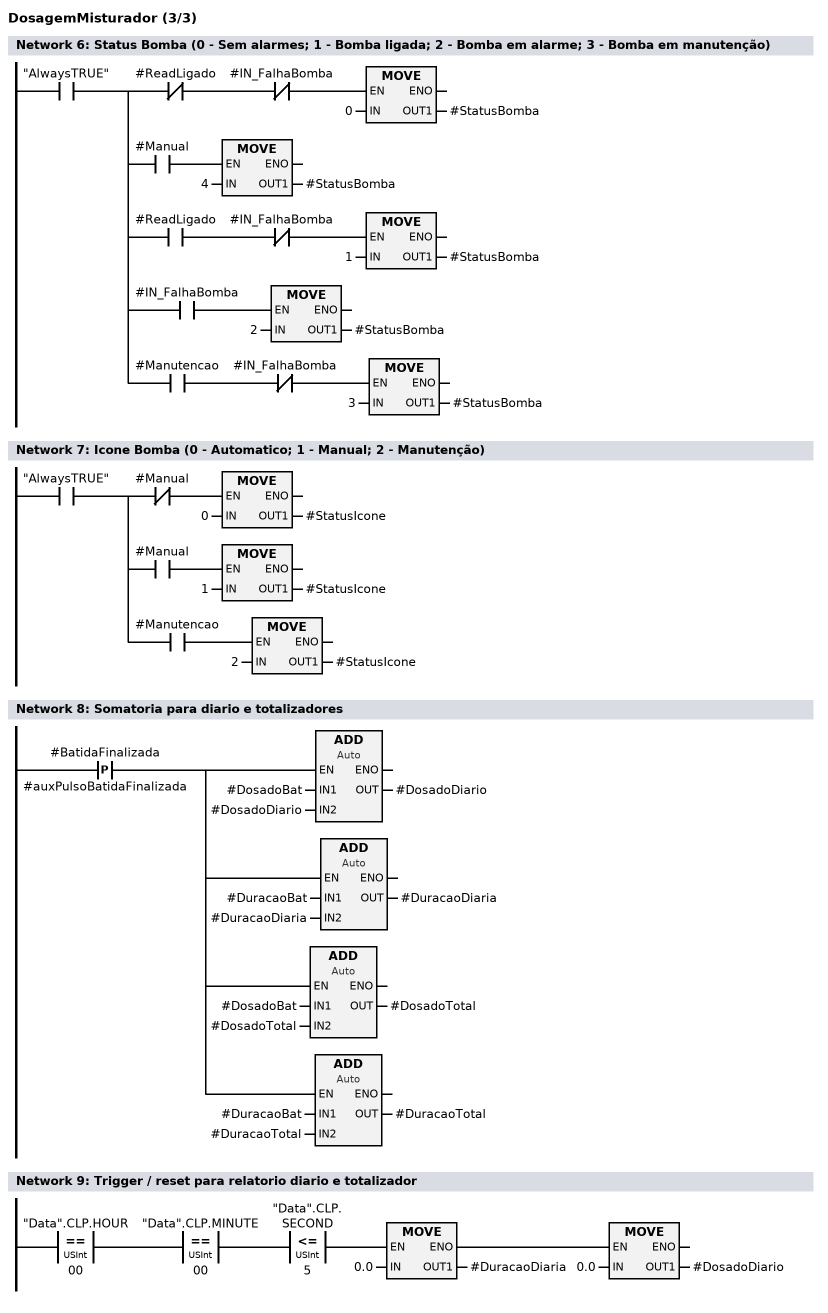
   RUNG wire#powerrail
      Contact( "AlwaysTRUE" )
      wire#w1
      I_Contact( #ReadLigado )
      I_Contact( #IN_FalhaBomba )
      Move(in := 0, out1 => #StatusBomba)
   END_RUNG
   RUNG wire#w1
      Contact( #Manual )
      Move(in := 4, out1 => #StatusBomba)
   END_RUNG
   RUNG wire#w1
      Contact( #ReadLigado )
      I_Contact( #IN_FalhaBomba )
      Move(in := 1, out1 => #StatusBomba)
   END_RUNG
   RUNG wire#w1
      Contact( #IN_FalhaBomba )
      Move(in := 2, out1 => #StatusBomba)
   END_RUNG
   RUNG wire#w1
      Contact( #Manutencao )
      I_Contact( #IN_FalhaBomba )
      Move(in := 3, out1 => #StatusBomba)
   END_RUNG
   // the same network as SCL:
   IF "AlwaysTRUE" AND NOT #ReadLigado AND NOT #IN_FalhaBomba THEN #StatusBomba := 0; END_IF;
   IF "AlwaysTRUE" AND #Manual THEN #StatusBomba := 4; END_IF;
   IF "AlwaysTRUE" AND #ReadLigado AND NOT #IN_FalhaBomba THEN #StatusBomba := 1; END_IF;
   IF "AlwaysTRUE" AND #IN_FalhaBomba THEN #StatusBomba := 2; END_IF;
   IF "AlwaysTRUE" AND #Manutencao AND NOT #IN_FalhaBomba THEN #StatusBomba := 3; END_IF;
END_REGION

REGION Network 7: Icone Bomba (0 - Automatico; 1 - Manual; 2 - Manutenção)
   RUNG wire#powerrail
      Contact( "AlwaysTRUE" )
      wire#w1
      I_Contact( #Manual )
      Move(in := 0, out1 => #StatusIcone)
   END_RUNG
   RUNG wire#w1
      Contact( #Manual )
      Move(in := 1, out1 => #StatusIcone)
   END_RUNG
   RUNG wire#w1
      Contact( #Manutencao )
      Move(in := 2, out1 => #StatusIcone)
   END_RUNG
   // the same network as SCL:
   IF "AlwaysTRUE" AND NOT #Manual THEN #StatusIcone := 0; END_IF;
   IF "AlwaysTRUE" AND #Manual THEN #StatusIcone := 1; END_IF;
   IF "AlwaysTRUE" AND #Manutencao THEN #StatusIcone := 2; END_IF;
END_REGION

REGION Network 8: Somatoria para diario e totalizadores
   RUNG wire#powerrail
      P_Contact(operand := #BatidaFinalizada, bit := #auxPulsoBatidaFinalizada)
      wire#w1
      Add(in1 := #DosadoBat, in2 := #DosadoDiario, out => #DosadoDiario)
   END_RUNG
   RUNG wire#w1
      Add(in1 := #DuracaoBat, in2 := #DuracaoDiaria, out => #DuracaoDiaria)
   END_RUNG
   RUNG wire#w1
      Add(in1 := #DosadoBat, in2 := #DosadoTotal, out => #DosadoTotal)
   END_RUNG
   RUNG wire#w1
      Add(in1 := #DuracaoBat, in2 := #DuracaoTotal, out => #DuracaoTotal)
   END_RUNG
   // the same network as SCL:
   #_w1 := #BatidaFinalizada AND NOT #auxPulsoBatidaFinalizada;   // rising edge of #BatidaFinalizada
   #auxPulsoBatidaFinalizada := #BatidaFinalizada;
   IF #_w1 THEN
       #DosadoDiario := #DosadoBat + #DosadoDiario;
       #DuracaoDiaria := #DuracaoBat + #DuracaoDiaria;
       #DosadoTotal := #DosadoBat + #DosadoTotal;
       #DuracaoTotal := #DuracaoBat + #DuracaoTotal;
   END_IF;
END_REGION

REGION Network 9: Trigger / reset para relatorio diario e totalizador
   RUNG wire#powerrail
      { S7_Templates := "SrcType := USInt" } EQ_Contact(in1 := "Data".CLP.HOUR, in2 := 00)
      { S7_Templates := "SrcType := USInt" } EQ_Contact(in1 := "Data".CLP.MINUTE, in2 := 00)
      { S7_Templates := "SrcType := USInt" } LE_Contact(in1 := "Data".CLP.SECOND, in2 := 5)
      Move(in := 0.0, out1 => #DuracaoDiaria)
      Move(in := 0.0, out1 => #DosadoDiario)
   END_RUNG
   // the same network as SCL:
   IF ("Data".CLP.HOUR = 00) AND ("Data".CLP.MINUTE = 00) AND ("Data".CLP.SECOND <= 5) THEN
       #DuracaoDiaria := 0.0;
       #DosadoDiario := 0.0;
   END_IF;
END_REGION
END_FUNCTION_BLOCK

FUNCTION_BLOCK "DosagemContinua"   // FB102, LAD
{ S7_Optimized_Access := 'TRUE' }
VERSION : 0.1
   VAR_INPUT
      SistemaHabilitado : Bool;
      Emergencia : Bool;
      SinalDosagem : Bool;
      PulsoMedidor : Bool;
      VolumePulso_ml : Real := 1.0;
      RetLigado : Bool;
      RetValvula : Bool;
      SP_DelayFinal : Time;
      SP_Dosagem : Real;
      VazaoNominalBBA : Real;
      IN_FalhaBomba : Bool;
      MedidorEstragado : Bool;
   END_VAR
   VAR_OUTPUT
      LigarValvula : Bool;
      LigarBomba : Bool;
      PorcentSaida : Real;
   END_VAR
   VAR RETAIN
      TON_DelayValvula : TON_TIME;
      Manual : Bool;
      LigaManual : Bool;
      Manutencao : Bool;
      StatusBomba : Int;
      StatusIcone : Int;
      TON_DelayAcionamento : TON_TIME;
      auxLigarValvula : Bool;
      TOF_RetardoValvula : TOF_TIME;
      TOF_RetardoDosagem : TOF_TIME;
      FatorAjuste : Real;
      VolumeAcionamento : Real;
      pPulsoMedidor : Bool;
      pClock10Hz : Bool;
      DuracaoAcionamento : Real;
      nLigarBomba : Bool;
      ResetFatorAjuste : Bool;
      DosagemAlvo : Real;
      auxDelayFinal : DInt;
      TON_ZeraAcumulados : TON_TIME;
      TOF_CalculaFator : TOF_TIME;
   END_VAR
   VAR_TEMP   // added for the SCL form of the ladder/FBD networks
      _w1 : Bool;
      _w2 : Bool;
      _w3 : Bool;
      _w4 : Bool;
   END_VAR
BEGIN

REGION Network 1: Dosa em automatico e manual
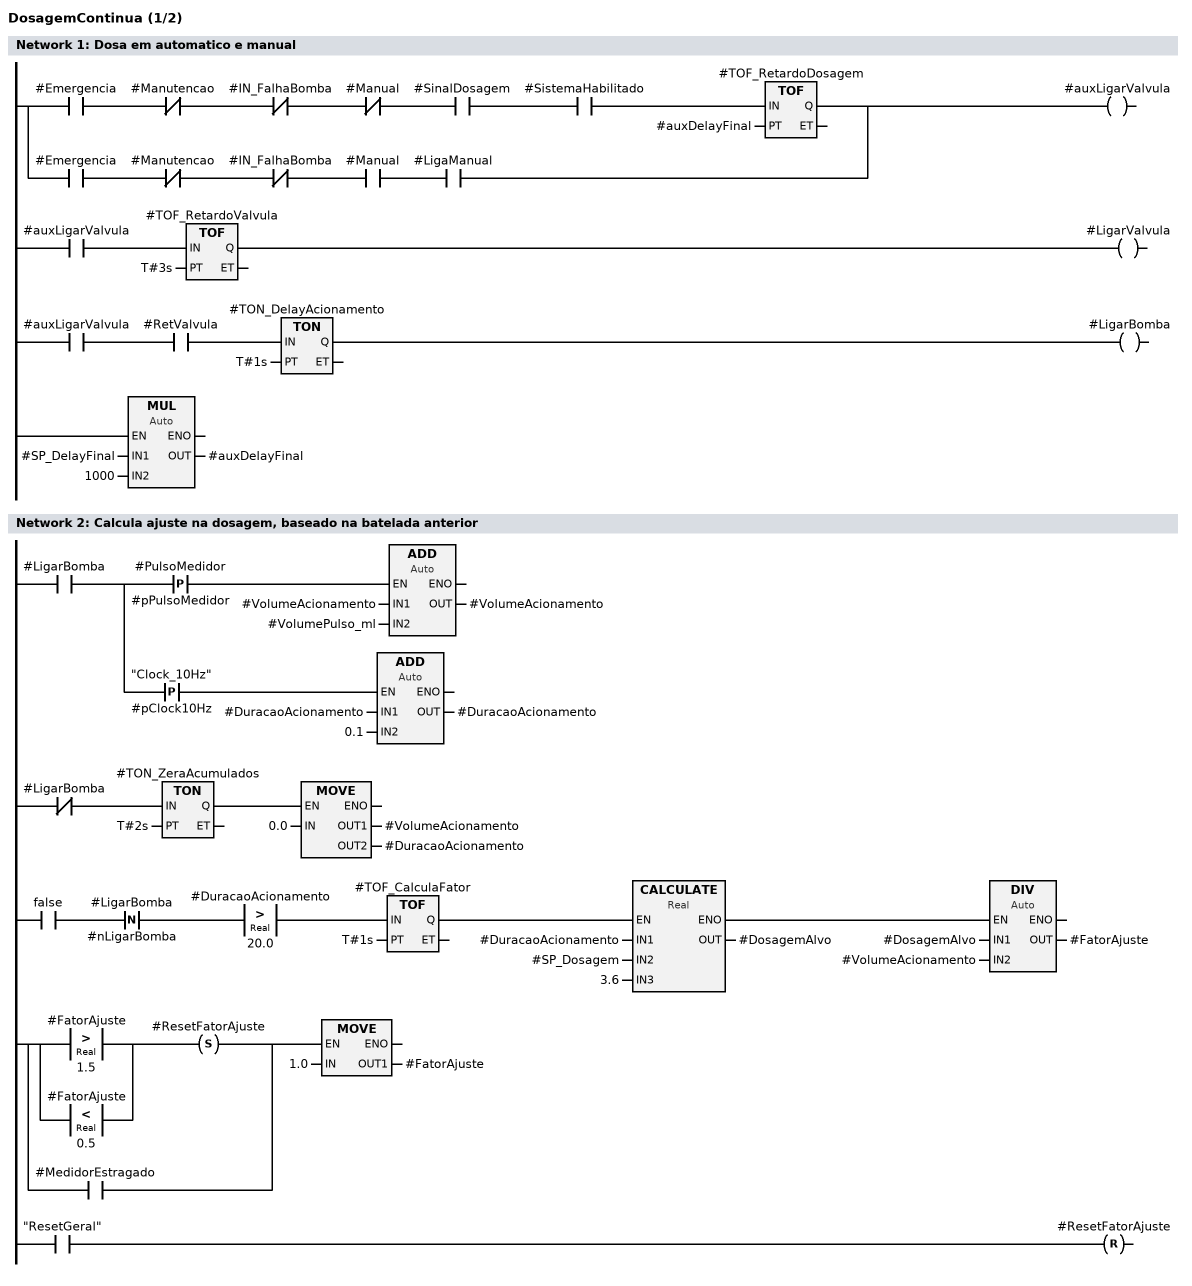
   #TOF_RetardoDosagem(IN := #Emergencia AND NOT #Manutencao AND NOT #IN_FalhaBomba AND NOT #Manual AND #SinalDosagem AND #SistemaHabilitado,   // TOF
                       PT := #auxDelayFinal);
   #auxLigarValvula := #TOF_RetardoDosagem.Q OR (#Emergencia AND NOT #Manutencao AND NOT #IN_FalhaBomba AND #Manual AND #LigaManual);
   #TOF_RetardoValvula(IN := #auxLigarValvula, PT := T#3s);   // TOF
   #LigarValvula := #TOF_RetardoValvula.Q;
   #TON_DelayAcionamento(IN := #auxLigarValvula AND #RetValvula, PT := T#1s);   // TON
   #LigarBomba := #TON_DelayAcionamento.Q;
   #auxDelayFinal := #SP_DelayFinal * 1000;
END_REGION

REGION Network 2: Calcula ajuste na dosagem, baseado na batelada anterior
   #_w1 := #LigarBomba AND #PulsoMedidor AND NOT #pPulsoMedidor;   // rising edge of #PulsoMedidor
   #pPulsoMedidor := #PulsoMedidor;
   IF #_w1 THEN #VolumeAcionamento := #VolumeAcionamento + #VolumePulso_ml; END_IF;
   #_w2 := #LigarBomba AND "Clock_10Hz" AND NOT #pClock10Hz;   // rising edge of "Clock_10Hz"
   #pClock10Hz := "Clock_10Hz";
   IF #_w2 THEN #DuracaoAcionamento := #DuracaoAcionamento + 0.1; END_IF;
   #TON_ZeraAcumulados(IN := NOT #LigarBomba, PT := T#2s);   // TON
   IF #TON_ZeraAcumulados.Q THEN
       #VolumeAcionamento := 0.0;
       #DuracaoAcionamento := 0.0;
   END_IF;
   #_w3 := false AND NOT #LigarBomba AND #nLigarBomba;   // falling edge of #LigarBomba
   #nLigarBomba := #LigarBomba;
   #TOF_CalculaFator(IN := #_w3 AND (#DuracaoAcionamento > 20.0), PT := T#1s);   // TOF
   IF #TOF_CalculaFator.Q THEN
       #DosagemAlvo := (#DuracaoAcionamento * #SP_Dosagem / 3.6);
       #FatorAjuste := #DosagemAlvo / #VolumeAcionamento;
   END_IF;
   #_w4 := (#FatorAjuste > 1.5) OR (#FatorAjuste < 0.5);
   IF #_w4 THEN #ResetFatorAjuste := TRUE; END_IF;
   IF #_w4 OR #MedidorEstragado THEN #FatorAjuste := 1.0; END_IF;
   IF "ResetGeral" THEN #ResetFatorAjuste := FALSE; END_IF;
END_REGION

REGION Network 3: Define % de dosagem da bomba
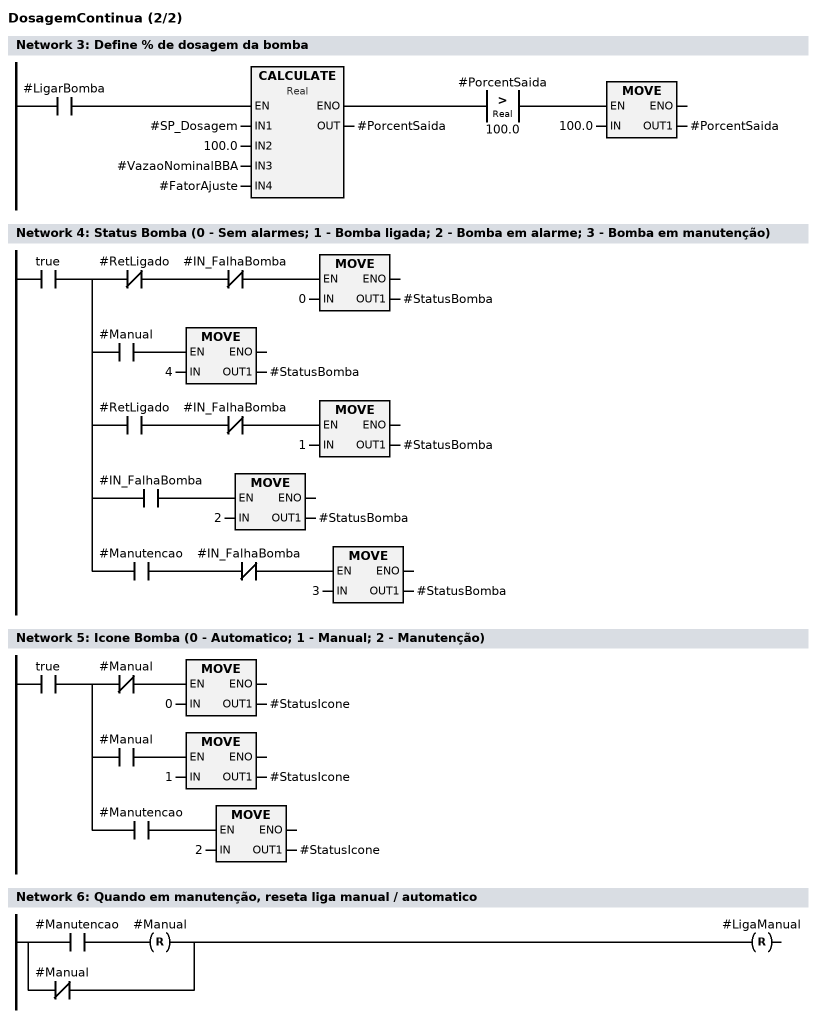
   RUNG wire#powerrail
      Contact( #LigarBomba )
      { S7_Templates := "SrcType := Real"; S7_Expression := "((IN1 * IN2 / IN3) * IN4)" } Calculate(in1 := #SP_Dosagem, in2 := 100.0, in3 := #VazaoNominalBBA, in4 := #FatorAjuste, out => #PorcentSaida)
      { S7_Templates := "SrcType := Real" } GT_Contact(in1 := #PorcentSaida, in2 := 100.0)
      Move(in := 100.0, out1 => #PorcentSaida)
   END_RUNG
   // the same network as SCL:
   IF #LigarBomba THEN #PorcentSaida := ((#SP_Dosagem * 100.0 / #VazaoNominalBBA) * #FatorAjuste); END_IF;
   IF #LigarBomba AND (#PorcentSaida > 100.0) THEN #PorcentSaida := 100.0; END_IF;
END_REGION

REGION Network 4: Status Bomba (0 - Sem alarmes; 1 - Bomba ligada; 2 - Bomba em alarme; 3 - Bomba em manutenção)
   RUNG wire#powerrail
      Contact( true )
      wire#w1
      I_Contact( #RetLigado )
      I_Contact( #IN_FalhaBomba )
      Move(in := 0, out1 => #StatusBomba)
   END_RUNG
   RUNG wire#w1
      Contact( #Manual )
      Move(in := 4, out1 => #StatusBomba)
   END_RUNG
   RUNG wire#w1
      Contact( #RetLigado )
      I_Contact( #IN_FalhaBomba )
      Move(in := 1, out1 => #StatusBomba)
   END_RUNG
   RUNG wire#w1
      Contact( #IN_FalhaBomba )
      Move(in := 2, out1 => #StatusBomba)
   END_RUNG
   RUNG wire#w1
      Contact( #Manutencao )
      I_Contact( #IN_FalhaBomba )
      Move(in := 3, out1 => #StatusBomba)
   END_RUNG
   // the same network as SCL:
   IF true AND NOT #RetLigado AND NOT #IN_FalhaBomba THEN #StatusBomba := 0; END_IF;
   IF true AND #Manual THEN #StatusBomba := 4; END_IF;
   IF true AND #RetLigado AND NOT #IN_FalhaBomba THEN #StatusBomba := 1; END_IF;
   IF true AND #IN_FalhaBomba THEN #StatusBomba := 2; END_IF;
   IF true AND #Manutencao AND NOT #IN_FalhaBomba THEN #StatusBomba := 3; END_IF;
END_REGION

REGION Network 5: Icone Bomba (0 - Automatico; 1 - Manual; 2 - Manutenção)
   RUNG wire#powerrail
      Contact( true )
      wire#w1
      I_Contact( #Manual )
      Move(in := 0, out1 => #StatusIcone)
   END_RUNG
   RUNG wire#w1
      Contact( #Manual )
      Move(in := 1, out1 => #StatusIcone)
   END_RUNG
   RUNG wire#w1
      Contact( #Manutencao )
      Move(in := 2, out1 => #StatusIcone)
   END_RUNG
   // the same network as SCL:
   IF true AND NOT #Manual THEN #StatusIcone := 0; END_IF;
   IF true AND #Manual THEN #StatusIcone := 1; END_IF;
   IF true AND #Manutencao THEN #StatusIcone := 2; END_IF;
END_REGION

REGION Network 6: Quando em manutenção, reseta liga manual / automatico
   RUNG wire#powerrail
      Contact( #Manutencao )
      R_Coil( #Manual )
      wire#w1
      R_Coil( #LigaManual )
   END_RUNG
   RUNG wire#powerrail
      I_Contact( #Manual )
   END_RUNG wire#w1
   // the same network as SCL:
   IF #Manutencao THEN #Manual := FALSE; END_IF;
   IF #Manutencao OR NOT #Manual THEN #LigaManual := FALSE; END_IF;
END_REGION
END_FUNCTION_BLOCK

FUNCTION_BLOCK "FBGammaX_1200"   // FB104, SCL
TITLE = Profibus GammaX
{ S7_Optimized_Access := 'TRUE' }
AUTHOR : kellerc
FAMILY : GammaX
NAME : Basic
VERSION : 1.0
// Erstellungsdatum:
// 
// Funktionsbeschreibung:
// 
// Änderungen:
   VAR_INPUT
      I_Adr_Status : Int;   // Adresse Int Eingang Steckplatz 1 DP-Kennung GammaX
      I_Adr_Operation_Mode : Int;   // Adresse Int Eingang Steckplatz 3 DP-Kennung GammaX
      I_Adr_Discharge : Int;   // Adresse Int Eingang Steckplatz 4 DP-Kennung GammaX
      I_Adr_Maximum_Discharge : Int;   // Adresse Int Eingang Steckplatz 5 DP-Kennung GammaX
      I_Adr_Batch : Int;   // Adresse Int Eingang Steckplatz 6 DP-Kennung GammaX
      I_Adr_Concentration : Int;   // Adresse Int Eingang Steckplatz 8 DP-Kennung GammaX
      I_Adr_Error_Warning : Int;   // Adresse Int Eingang Steckplatz 10 DP-Kennung GammaX
      I_Adr_Stroke_Quantity : Int;   // Adresse Int Eingang Steckplatz 11 DP-Kennung GammaX
      O_Adr_Control : Int;   // Adresse Int Ausgang Steckplatz 2 DP-Kennung GammaX
      O_Adr_Operation_Mode : Int;   // Adresse Int Ausgang Steckplatz 3 DP-Kennung GammaX
      O_Adr_Discharge : Int;   // Adresse Int Ausgang Steckplatz 4 DP-Kennung GammaX
      O_Adr_Batch : Int;   // Adresse Int Ausgang Steckplatz 6 DP-Kennung GammaX
      O_Adr_Contact : Int;   // Adresse Int Ausgang Steckplatz 7 DP-Kennung GammaX
      O_Adr_Concentration : Int;   // Adresse Int Ausgang Steckplatz 8 DP-Kennung GammaX
      O_Adr_Metering_Monitor : Int;   // Adresse Int Ausgang Steckplatz 9 DP-Kennung GammaX
      O_Adr_Stroke_Quantity : Int;   // Adresse Int Ausgang Steckplatz 11 DP-Kennung GammaX
      ixStart_Stop : Bool;   // Eingang Start/Stop 0=Stopp 1=Start
      ixStartBatch_Or_Contact : Bool;   // Eingang Wenn sich der Wert von 0 auf 1 ändert, wird im Chargenbetrieb eine Char
      ixBatchContactMemory : Bool;   // Eingang Ist der Chargenspeicher aktiviert und wird während einer laufenden Char
      ixMeteringMonitor : Bool;   // Bei installierter Dosierüberwachung kann sie selbst eingeschaltet werden (1). A
      ixReset : Bool;   // Eingang Reset 0 -> 1 Flanke führt Reset aus
      ixResetPump : Bool;   // Wenn der Wert von Reset von 1 auf 0 wechselt, wird der interne Pumpenspeicher g
      ixFault_Lock : Bool;   // Eingang Verriegelung bei Fehler 0=keine Verriegelung bei Fehler, 1=Verriegelung
      ixResetStrokeCounter : Bool;   // Eingang Reset Hubzähler, Reset bei 0 -> 1 Flanke
      ixResetQuantity : Bool;   // Eingang Reset Mengenzähler, Reset bei 0 -> 1 Flanke
      ixFlowControl_OnOff : Bool;   // Eingang Bei installierter Dosierüberwachung, kann sie eingeschaltet ( 1) werden
      ixModeSetpoint : Bool;   // 0 = 0-100%, 1 = Liter pro Stunde
      iyMode : Byte;   // Eingang Modus der Pumpe 0=Aus,1=Manual,2=Batch,3=Kontakt,4=Analog,17=(Konz),18=
      irSetpoint_0_100 : Real;   // Eingang Sollwert Dosierpumpe 0-100%
      irSetpoint_Volume : Real;   // Eingang Sollwert Dosierpumpe als Volume
      irBatchVolume : Real;   // Dosiervolumen einer Charge
      iiBatchTime : Int;   // Zeit, in welcher Charge dosiert werden soll
      irContactVolume : Real;   // Dosiervolumen, das pro Kontakt dosiert werden soll
      irConcentration : Real;   // Sollwert der Konzentrationseinstellung (nur bei Betriebsart Konzentation)
      iiCycle_Error : Int;   // Anzahl Zyklen bis Fehler angezeigt wird
   END_VAR
   VAR_OUTPUT
      oxRunning : Bool;   // Ausgang Dosierpumpe läuft 0=läuft nicht 1=läuft
      oxWarning : Bool;   // Ausgang Warnung Dosierpumpe 0=keine Warnung 1=Warnung
      oxError : Bool;   // Ausgang Störung Dosierpumpe 0=keine Störung 1=Störung
      oxWarningProfibus : Bool;   // Ausgang Störung Profibus 0=keine Warnung 1=Warnung (Pumpe nicht steuerbar)
      oyMode : Byte;   // Eingang Modus der Pumpe 0=Aus,1=Manual,2=Batch,3=Kontakt,4=Analog,17=(Konz),18=
      orFlowrate : Real;   // Istwert Dosierleistung
      orMaxFlowrate : Real;   // Maximale Dosierleistung in l/h
      orConcentration : Real;   // Ausgang Ist an der Pumpe die Konzentrationsberechnung aktiviert, kann die aktue
      orRemainingVolumeInBatch : Real;   // noch zu dosierendes Restvolumen beim Batchbetrieb
      odStrokeCounter : DInt;   // Ausgang Hubzähler
      orQuantityCounter : Real;   // Ausgang Mengenzähler in Liter
      orLitersPerStroke : Real;   // Liter pro Hub
   END_VAR
   VAR
      Status : Struct
         Service : Bool;   // 1=Es sind Serviceanforderungen vorhanden, 0= Es sind keine Serviceanforderungen
         Messages : Bool;   // 1=Es sind Meldungen vorhanden, 0=Es sind keine Meldungen vorhanden
         Error : Bool;   // 1=Störung, 0=keine Störung
         Warnings : Bool;   // 1=Warnung, 0=keine Warnung
         ManuelStop : Bool;   // 1=Pumpe wurde von Hand gestoppt, 0=Pumpe ist nicht von Hand gestoppt
         Stop : Bool;   // 1=Pumpe ist gestoppt, 0=Pumpe ist nicht gestoppt
         Intake : Bool;   // 1=Ansaugen aktiv, 0=Ansaugen inaktiv
         Auxiliary : Bool;   // 1=Pumpe ist in Auxiliarbetrieb, 0=Pumpe ist nicht in Auxiliarbetrieb
         Pause : Bool;   // 1=Pause aktiv, 0=Pause inaktiv
         Module : Bool;   // 0=kein Profibus aktiviert, oder Profibus gestört -> Pumpe nicht steuerbar 1=Pro
         Flow : Bool;   // 0=Dosierüberwachung inaktiv, 1=Dosierüberwachung aktiv
         BatchMemory : Bool;   // 0=Batch Speicher ist nicht aktiviert, 1=Batch Speicher aktiviert
         Calibrated : Bool;   // 0=Pumpe ist nicht kalibriert, 1=Pumpe ist kalibriert
         NotUsed1 : Bool;   // nicht benutzt
         NotUsed2 : Bool;   // nicht benutzt
         NotUsed3 : Bool;   // nicht benutzt
         Diaphragm : Bool;   // 0=Membranbruchsensor nicht vorhanden, 1=Membranbruchsensor vorhanden
         Concentration : Bool;   // 0=Konzentrationsberechnung nicht aktiv, 1=Konzentrationsberechnung aktiv
         NotUsed4 : Bool;   // nicht benutzt
         Overpressure : Bool;   // 0=OK, 1=Antriebssteuerung meldet zu hoher Gegendruck
         Depressurised : Bool;   // 0=OK, 1=Antriebssteuerung meldet kein Gegendruck
         Venting : Bool;   // 0=OK, 1=Pumpe entlüftet im Moment
         NotUsed5 : Bool;   // nicht benutzt
         NotUsed6 : Bool;   // nicht benutzt
         NotUsed7 : Bool;   // nicht benutzt
         NotUsed8 : Bool;   // nicht benutzt
         NotUsed9 : Bool;   // nicht benutzt
      END_STRUCT;
      Errors : Struct
         Minimum : Bool;   // 0 = kein Fehler, 1 = Dosierflüssigkeitsstand zu gering
         Batch : Bool;   // 0 = kein Fehler, 1 = Zu viele Dosierhübe > 100000
         Analog_4mA : Bool;   // 0 = kein Fehler, 1 = Analogstrom ist kleiner 4 mA
         Analog_20mA : Bool;   // 0 = kein Fehler, 1 = Analogstrom ist größer 23 mA
         FlowMonitoring : Bool;   // 0 = kein Fehler, 1 = Dosierüberwachungsfehler
         DiaphragmFailure : Bool;   // 0 = kein Fehler, 1 = Defekte Membran im Dosierkopf
         AirLock : Bool;   // 0 = kein Fehler, 1 = Luft im Dosierkopf
         Overpressure : Bool;   // 0 = kein Fehler, 1 = Überdruck in der Hydraulik
         NotUsed1 : Bool;   // nicht benutzt
         Cavitation : Bool;   // 0 = kein Fehler, 1 = Kaviatation
         LowPressure : Bool;   // 0 = kein Fehler, 1 = Zu geringer Druck in der Hydraulik
         StrokeLenghtChanged : Bool;   // 0 = kein Fehler, 1 = Im gesperrten Zustand wurde die Hublänge geändert
         Venting : Bool;   // 0 = kein Fehler, 1 = Automatische Entlüftung nicht möglich
         BusError : Bool;   // 0 = kein Fehler, 1 = Vom Modul gemeldeter Busfehler
         SystemError : Bool;   // 0 = kein Fehler, 1 = Systemkomponenten defekt. Siehe Display
         ModuleError : Bool;   // 0 = kein Fehler, 1 = Fehler im Modulhandling
      END_STRUCT;
      Warnings : Struct
         Minimum : Bool;   // 0 = keine Warnung, 1 = Dosierflüssigkeitsstand ist gering
         Calibration : Bool;   // 0 = keine Warnung, 1 = Hublängeneinstellung außerhalb der Kalibriertoleranz
         FlowMonitoring : Bool;   // 0 = keine Warnung, 1 = Dosierüberwachungswarnung
         DiaphragmFailure : Bool;   // 0 = keine Warnung, 1 = Defekte Membran im Dosierkopf
         Airlock : Bool;   // 0 = keine Warnung, 1 = Luft im Dosierkopf
         NotUsed1 : Bool;   // nicht benutzt
         Cavitation : Bool;   // 0 = keine Warnung, 1 = Kaviatation
         Overpressure : Bool;   // 0 = keine Warnung, 1 = Überdruck in der Hydraulik
         LowPressure : Bool;   // 0 = keine Warnung, 1 = Zu geringer Druck in der Hydraulik
      END_STRUCT;
      iiCycleFault : Int;
      iiCycleWarning : Int;
   END_VAR
   VAR_TEMP
      temp_Setpoint : Real;   // Temporärer Setpoint der Pumpe
      temp_byte : Byte;   // Temporärer Byte für Perepheriezugriffe
      temp_word : Word;
      temp_int : Int;
      temp_byte2 : Byte;
      temp_dword : DWord;
      temp_status_0 : Byte;
      temp_status_1 : Byte;
      temp_status_2 : Byte;
      temp_status_3 : Byte;
      temp_Error_0 : Byte;
      temp_Error_1 : Byte;
      temp_Warning_0 : Byte;
      temp_Warning_1 : Byte;
   END_VAR
BEGIN

   (*
               #temp_byte := 16#01;
               POKE(area := 16#82,
                   dbNumber := 0,
                   byteOffset := #O_Adr_Control,
                   value := #temp_byte);



   PEEK_WORD(area := 16#81, dbNumber := 0, byteOffset := #I_Adr_Max_Frequency);                
   PEEK_DWORD(area := 16#81, dbNumber := 0, byteOffset := #I_Adr_Max_Frequency);                
   *)




       // Anweisungsteil
       #orFlowrate := DWORD_TO_REAL(PEEK_DWORD(area := 16#81, dbNumber := 0, byteOffset := #I_Adr_Discharge));//%ED(#I_Adr_Discharge):P);
       #orMaxFlowrate := DWORD_TO_REAL(PEEK_DWORD(area := 16#81, dbNumber := 0, byteOffset := #I_Adr_Maximum_Discharge));//%ED(#I_Adr_Maximum_Discharge):P);    


       IF #ixModeSetpoint = FALSE THEN
           #temp_Setpoint := #orMaxFlowrate * #irSetpoint_0_100 / 100.0;
       ELSE
           #temp_Setpoint := #irSetpoint_Volume;
       END_IF;


       IF #temp_Setpoint >= #orMaxFlowrate THEN
           #temp_Setpoint := #orMaxFlowrate;
       ELSIF #temp_Setpoint <= 0.0 THEN
           #temp_Setpoint := 0.0;
       END_IF;



       #temp_dword := REAL_TO_DWORD(#temp_Setpoint );
       POKE(area := 16#82,
            dbNumber := 0,
            byteOffset := #O_Adr_Discharge,
            value := #temp_dword);
       // %AD(#O_Adr_Discharge):P := REAL_TO_DWORD(#temp_Setpoint );


       POKE(area := 16#82,
            dbNumber := 0,
            byteOffset := #O_Adr_Operation_Mode,
            value := #iyMode);
       //%AB(#O_Adr_Operation_Mode):P := #iyMode;

       IF #ixStart_Stop = true THEN
           #temp_byte2 := 16#01;
           POKE(area := 16#82,
                dbNumber := 0,
                byteOffset := #O_Adr_Control,
                value := #temp_byte2);
           //%AB(#O_Adr_Control):P := 16#01;
       ELSE
           #temp_byte2 := 16#00;
           POKE(area := 16#82,
                dbNumber := 0,
                byteOffset := #O_Adr_Control,
                value := #temp_byte2);
           //%AB(#O_Adr_Control):P := 16#00;
       END_IF;


       IF #ixResetPump = false THEN
           #temp_byte2 := 16#00;
           POKE(area := 16#82,
                dbNumber := 0,
                byteOffset := #O_Adr_Control + 1,
                value := #temp_byte2);
           //%AB(#O_Adr_Control + 1):P := 16#00;
       ELSE
           #temp_byte2 := 16#00;
           POKE(area := 16#82,
                dbNumber := 0,
                byteOffset := #O_Adr_Control + 1,
                value := #temp_byte2);
           //%AB(#O_Adr_Control + 1):P := 16#01;
       END_IF;



       // Status Ausgang


           IF #orFlowrate > 0.0 THEN
               #oxRunning := true;
           ELSE
               #oxRunning := false;
           END_IF;



           // Status Mode
           //#temp_byte := SHR (IN := %EB(#I_Adr_Status+3):P, N := 2) AND 16#07; // TODO: Wird diese Auswertung entfernt? Oder wird PEB[I_Adr_Operation_Mode] genutzt
           #oyMode := PEEK_BYTE(area := 16#81, dbNumber := 0, byteOffset := #I_Adr_Operation_Mode); //%EB(#I_Adr_Operation_Mode):P;

           #temp_status_0 := PEEK_BYTE(area := 16#81, dbNumber := 0, byteOffset := #I_Adr_Status);
           #temp_status_1 := PEEK_BYTE(area := 16#81, dbNumber := 0, byteOffset := #I_Adr_Status + 1);
           #temp_status_2 := PEEK_BYTE(area := 16#81, dbNumber := 0, byteOffset := #I_Adr_Status + 2);
           #temp_status_3 := PEEK_BYTE(area := 16#81, dbNumber := 0, byteOffset := #I_Adr_Status+ 3);


       // Status statischer Bereich
           #Status.Service := (#temp_status_3 AND 16#01) = 16#01;                                // 1=Service anstehend, 0=keine Service anstehend
           #Status.Messages := (#temp_status_3 AND 16#02) = 16#02;                                // 1=Meldung, 0=keine Meldung
           #Status.Error := (#temp_status_3 AND 16#20) = 16#20;                                // 1=Störung, 0=keine Störung
           #Status.Warnings := (#temp_status_3 AND 16#40) = 16#40;                                // 1=Warnung, 0=keine Warnung
           #Status.ManuelStop := (#temp_status_3 AND 16#80) = 16#80;                            // 1=Pumpe wurde von Hand gestoppt, 0=Pumpe ist nicht von Hand gestoppt
           #Status.Stop := (#temp_status_2 AND 16#01) = 16#01;                                 // 1=Pumpe ist gestoppt, 0=Pumpe ist nicht gestoppt
           #Status.Intake := (#temp_status_2 AND 16#02) = 16#02;                               // 1=Ansaugen aktiv, 0=Ansaugen inaktiv
           #Status.Auxiliary :=(#temp_status_2 AND 16#04) = 16#04;                             // 1=Pumpe ist in Auxiliarbetrieb, 0=Pumpe ist nicht in Auxiliarbetrieb
           #Status.Pause := (#temp_status_2 AND 16#08) = 16#08;                                // 1=Pause aktiv, 0=Pause inaktiv
           #Status.Module := (#temp_status_2 AND 16#10) = 16#10;                               // 0=Automatic Mode???
           #Status.Flow := (#temp_status_2 AND 16#20) = 16#20;                                 // 0=Dosierüberwachung inaktiv, 1=Dosierüberwachung aktiv
           #Status.BatchMemory := (#temp_status_2 AND 16#40)= 16#40;                           // 0=Batch Speicher ist nicht aktiviert, 1=Batch Speicher aktiviert
           #Status.Calibrated := (#temp_status_2 AND 16#80) = 16#80;                           // 0=Pumpe ist nicht kalibriert, 1=Pumpe ist kalibriert
           #Status.NotUsed1 := (#temp_status_1 AND 16#01) = 16#01;                             // nicht benutzt
           #Status.NotUsed2 := (#temp_status_1 AND 16#02) = 16#02;                             // nicht benutzt
           #Status.NotUsed3 := (#temp_status_1 AND 16#04) = 16#04;                                // nicht benutzt
           #Status.Diaphragm := (#temp_status_1 AND 16#08) = 16#08;                            // 0=Membranbruchsensor nicht vorhanden, 1=Membranbruchsensor vorhanden
           #Status.Concentration := (#temp_status_1 AND 16#10) = 16#10;                        // 0=Konzentrationsberechnung nicht aktiv, 1=Konzentrationsberechnung aktiv
           #Status.NotUsed4 := (#temp_status_1 AND 16#80) = 16#80;                             // nicht benutzt
           #Status.Overpressure := (#temp_status_0 AND 16#01) = 16#01;                           // 0=OK, 1=Antriebssteuerung meldet zu hoher Gegendruck
           #Status.Depressurised := (#temp_status_0 AND 16#02) = 16#02;                          // 0=OK, 1=Antriebssteuerung meldet kein Gegendruck
           #Status.Venting := (#temp_status_0 AND 16#04) = 16#04;                                // 0=OK, 1=Pumpe entlüftet im Moment
           #Status.NotUsed5 := (#temp_status_0 AND 16#08) = 16#08;                               // nicht benutzt
           #Status.NotUsed6 := (#temp_status_0 AND 16#10) = 16#10;                                 // nicht benutzt
           #Status.NotUsed7 := (#temp_status_0 AND 16#20) = 16#20;                                // nicht benutzt
           #Status.NotUsed8 := (#temp_status_0 AND 16#40) = 16#40;                                // nicht benutzt
           #Status.NotUsed9 := (#temp_status_0 AND 16#80) = 16#80;                                // nicht benutzt
       // Ende Status statischer Bereich


           #temp_Error_0 := PEEK_BYTE(area := 16#81, dbNumber := 0, byteOffset := #I_Adr_Error_Warning + 3);
           #temp_Error_1 := PEEK_BYTE(area := 16#81, dbNumber := 0, byteOffset := #I_Adr_Error_Warning + 2);
           #temp_Warning_0 := PEEK_BYTE(area := 16#81, dbNumber := 0, byteOffset := #I_Adr_Error_Warning + 5);
           #temp_Warning_1 := PEEK_BYTE(area := 16#81, dbNumber := 0, byteOffset := #I_Adr_Error_Warning + 4);



       // Anfang Error statischer Bereich * Complete *
           #Errors.Minimum             := (#temp_Error_0 AND 16#01)  = 16#01;          // 0 = kein Fehler, 1 = Dosierflüssigkeitsstand zu gering
           #Errors.Batch               := (#temp_Error_0 AND 16#02)  = 16#02;          // 0 = kein Fehler, 1 = Zu viele Dosierhübe > 100000
           #Errors.Analog_4mA          := (#temp_Error_0 AND 16#04)  = 16#04;          // 0 = kein Fehler, 1 = Analogstrom ist kleiner 4 mA
           #Errors.Analog_20mA         := (#temp_Error_0 AND 16#08)  = 16#08;          // 0 = kein Fehler, 1 = Analogstrom ist größer 23 mA
           #Errors.FlowMonitoring      := (#temp_Error_0 AND 16#10)  = 16#10;          // 0 = kein Fehler, 1 = Dosierüberwachungsfehler
           #Errors.DiaphragmFailure    := (#temp_Error_0 AND 16#20)  = 16#20;          // 0 = kein Fehler, 1 = Defekte Membran im Dosierkopf
           #Errors.AirLock             := (#temp_Error_0 AND 16#40)  = 16#40;          // 0 = kein Fehler, 1 = Luft im Dosierkopf
           #Errors.Overpressure        := (#temp_Error_0 AND 16#80)  = 16#80;          // 0 = kein Fehler, 1 = Überdruck in der Hydraulik
           #Errors.NotUsed1            := (#temp_Error_1 AND 16#01)  = 16#01;            // nicht benutzt
           #Errors.Cavitation          := (#temp_Error_1 AND 16#02)  = 16#02;            // 0 = kein Fehler, 1 = Kaviatation        
           #Errors.LowPressure         := (#temp_Error_1 AND 16#04)  = 16#04;            // 0 = kein Fehler, 1 = Zu geringer Druck in der Hydraulik
           #Errors.StrokeLenghtChanged := (#temp_Error_1 AND 16#08)  = 16#08;          // 0 = kein Fehler, 1 = Im gesperrten Zustand wurde die Hublänge geändert
           #Errors.Venting             := (#temp_Error_1 AND 16#10)  = 16#10;          // 0 = kein Fehler, 1 = Automatische Entlüftung nicht möglich
           #Errors.BusError            := (#temp_Error_1 AND 16#20)  = 16#20;          // 0 = kein Fehler, 1 = Vom Modul gemeldeter Busfehler
           #Errors.SystemError         := (#temp_Error_1 AND 16#40)  = 16#40;          // 0 = kein Fehler, 1 = Systemkomponenten defekt. Siehe Display
           #Errors.ModuleError         := (#temp_Error_1 AND 16#80)  = 16#80;          // 0 = kein Fehler, 1 = Fehler im Modulhandling 
       // Ende Error statischer Bereich * Complete *

       // Anfang Warnings statischer Bereich * Complete *
           #Warnings.Minimum           := (#temp_Warning_0 AND 16#01)  = 16#01;          // 0 = keine Warnung, 1 = Dosierflüssigkeitsstand ist gering
           #Warnings.Calibration       := (#temp_Warning_0 AND 16#02)  = 16#02;          // 0 = keine Warnung, 1 = Hublängeneinstellung außerhalb der Kalibriertoleranz
           #Warnings.FlowMonitoring    := (#temp_Warning_0 AND 16#04)  = 16#04;          // 0 = keine Warnung, 1 = Dosierüberwachungswarnung
           #Warnings.DiaphragmFailure  := (#temp_Warning_0 AND 16#08)  = 16#08;          // 0 = keine Warnung, 1 = Defekte Membran im Dosierkopf
           #Warnings.Airlock           := (#temp_Warning_0 AND 16#10)  = 16#10;          // 0 = keine Warnung, 1 = Luft im Dosierkopf
           #Warnings.NotUsed1          := (#temp_Warning_0 AND 16#20)  = 16#20;            // nicht benutzt
           #Warnings.Cavitation        := (#temp_Warning_0 AND 16#40)  = 16#40;            // 0 = kein Fehler, 1 = Kaviatation
           #Warnings.Overpressure      := (#temp_Warning_0 AND 16#80)  = 16#80;          // 0 = keine Warnung, 1 = Überdruck in der Hydraulik
           #Warnings.LowPressure       := (#temp_Warning_1 AND 16#01)  = 16#01;          // 0 = keine Warnung, 1 = Zu geringer Druck in der Hydraulik
        // Ende Warnings statischer Bereich * Complete *   




   // Chargenbetrieb und Kontaktbetrieb
           IF #ixStartBatch_Or_Contact = TRUE THEN
               #temp_byte2 := 16#01;
               POKE(area := 16#82,
                    dbNumber := 0,
                    byteOffset := #O_Adr_Batch + 6,
                    value := #temp_byte2);
           //%AB(#O_Adr_Batch+5):P := 16#01;
           ELSE
               #temp_byte2 := 16#00;
               POKE(area := 16#82,
                    dbNumber := 0,
                    byteOffset := #O_Adr_Batch + 6,
                    value := #temp_byte2);
           //%AB(#O_Adr_Batch+5):P := 16#00;
       END_IF;

       IF #ixBatchContactMemory = TRUE THEN
           #temp_byte2 := 16#01;
           POKE(area := 16#82,
                dbNumber := 0,
                byteOffset := #O_Adr_Batch + 7,
                value := #temp_byte2);
           #temp_byte2 := 16#01;
           POKE(area := 16#82,
                dbNumber := 0,
                byteOffset := #O_Adr_Contact + 4,
                value := #temp_byte2);
           //%AB(#O_Adr_Batch+6):P := 16#01;
           //%AB(#O_Adr_Contact+4):P := 16#01;
       ELSE
           #temp_byte2 := 16#00;
           POKE(area := 16#82,
                dbNumber := 0,
                byteOffset := #O_Adr_Batch + 7,
                value := #temp_byte2);
           #temp_byte2 := 16#00;
           POKE(area := 16#82,
                dbNumber := 0,
                byteOffset := #O_Adr_Contact + 4,
                value := #temp_byte2);
           //%AB(#O_Adr_Batch+6):P := 16#00;
           //%AB(#O_Adr_Contact+4):P := 16#00;
       END_IF;

       #temp_dword := REAL_TO_DWORD(#irBatchVolume);
       POKE(area := 16#82,
            dbNumber := 0,
            byteOffset := #O_Adr_Batch,
            value := #temp_dword);
       //%AD(#O_Adr_Batch):P := REAL_TO_DWORD(#irBatchVolume);
       //
       #temp_word := INT_TO_WORD(#iiBatchTime);
       POKE(area := 16#82,
            dbNumber := 0,
            byteOffset := #O_Adr_Batch+4,
            value := #temp_word);
      // %AW(#O_Adr_Batch+4):P := INT_TO_WORD(#iiBatchTime);

       #temp_dword := REAL_TO_DWORD(#irContactVolume);
       POKE(area := 16#82,
            dbNumber := 0,
            byteOffset := #O_Adr_Contact,
            value := #temp_dword);
       //%AD(#O_Adr_Contact):P := REAL_TO_DWORD(#irContactVolume);

       #orRemainingVolumeInBatch := DWORD_TO_REAL(PEEK_DWORD(area := 16#81, dbNumber := 0, byteOffset := #I_Adr_Batch));//%ED(#I_Adr_Batch):P);
   // Chargenbetrieb und Kontaktbetrieb Ende

       #orConcentration := DWORD_TO_REAL(PEEK_DWORD(area := 16#81, dbNumber := 0, byteOffset := #I_Adr_Concentration));//%ED(#I_Adr_Concentration):P);

       #temp_dword := REAL_TO_DWORD(#irConcentration);
       POKE(area := 16#82,
            dbNumber := 0,
            byteOffset := #O_Adr_Concentration,
            value := #temp_dword);
       //%AD(#O_Adr_Concentration):P := REAL_TO_DWORD(#irConcentration);

       IF #ixMeteringMonitor = TRUE THEN
           #temp_byte2 := 16#01;
           POKE(area := 16#82,
                dbNumber := 0,
                byteOffset := #O_Adr_Metering_Monitor,
                value := #temp_byte2);
           //%AB(#O_Adr_Metering_Monitor):P := 16#01;
       ELSE
           #temp_byte2 := 16#00;
           POKE(area := 16#82,
                dbNumber := 0,
                byteOffset := #O_Adr_Metering_Monitor,
                value := #temp_byte2);
           //%AB(#O_Adr_Metering_Monitor):P := 16#00;
       END_IF;







   // Hubzähler Auslesen und Zurücksetzen      
       #odStrokeCounter := DWORD_TO_DINT(PEEK_DWORD(area := 16#81, dbNumber := 0, byteOffset := #I_Adr_Stroke_Quantity));//DWORD_TO_DINT(%ED(#I_Adr_Stroke_Quantity):P);

       IF #ixResetStrokeCounter = true THEN
           #temp_byte2 := 16#01;
           POKE(area := 16#82,
                dbNumber := 0,
                byteOffset := #O_Adr_Stroke_Quantity,
                value := #temp_byte2);
           //%AB(#O_Adr_Stroke_Quantity):P := 16#01;
       ELSE
           #temp_byte2 := 16#00;
           POKE(area := 16#82,
                dbNumber := 0,
                byteOffset := #O_Adr_Stroke_Quantity,
                value := #temp_byte2);
           //%AB(#O_Adr_Stroke_Quantity):P := 16#00;
       END_IF;

   // Mengenzähler Auslesen und Zurücksetzen      
       #orQuantityCounter := DWORD_TO_REAL(PEEK_DWORD(area := 16#81, dbNumber := 0, byteOffset := #I_Adr_Stroke_Quantity+4));//DWORD_TO_REAL(%ED(#I_Adr_Stroke_Quantity+4):P);

       IF #ixResetQuantity = true THEN
           #temp_byte2 := 16#01;
           POKE(area := 16#82,
                dbNumber := 0,
                byteOffset := #O_Adr_Stroke_Quantity+1,
                value := #temp_byte2);
           //%AB(#O_Adr_Stroke_Quantity+1):P := 16#01;
       ELSE
           #temp_byte2 := 16#00;
           POKE(area := 16#82,
                dbNumber := 0,
                byteOffset := #O_Adr_Stroke_Quantity + 1,
                value := #temp_byte2);
           //%AB(#O_Adr_Stroke_Quantity+1):P := 16#00;
       END_IF;

   // Hubmenge
       #orLitersPerStroke := DWORD_TO_REAL(PEEK_DWORD(area := 16#81, dbNumber := 0, byteOffset := #I_Adr_Stroke_Quantity+8));//DWORD_TO_REAL(%ED(#I_Adr_Stroke_Quantity+8):P);


       // Ende Status statischer Bereich

               IF #Status.Error = true AND #oxError = false THEN
               #iiCycleFault := #iiCycleFault + 1;
               IF #iiCycleFault >= #iiCycle_Error THEN
                   #oxError := true;
               END_IF;
           END_IF;

           IF #Status.Error = false AND #ixReset = true THEN
               #iiCycleFault := 0;
               #oxError := false;
           END_IF;

           IF #Status.Warnings = true AND #oxWarning = false THEN
               #iiCycleWarning := #iiCycleWarning + 1;
               IF #iiCycleWarning >= #iiCycle_Error THEN
                   #oxWarning := true;
               END_IF;
           END_IF;

           IF #Status.Warnings = false AND #ixReset = true THEN
               #iiCycleWarning := 0;
               #oxWarning := false;
           END_IF;  

           IF #Status.Module = false THEN
               #oxWarningProfibus := true;
           END_IF;

           IF #Status.Module = true AND #ixReset = true THEN
               #oxWarningProfibus := false;
           END_IF;
END_FUNCTION_BLOCK

// folder: FC

FUNCTION "FC_EspModbusCFW" : Void   // FC1, LAD
{ S7_Optimized_Access := 'TRUE' }
VERSION : 0.1
   VAR_IN_OUT
      ReadModbus : Array[1..7] of Int;
      WriteModbus : Array[0..1] of Int;
      Inversor : "ModbusCFW";
   END_VAR
BEGIN

REGION Network 1: 1 = Write Frequencia (hex) / 2 = Read Frequencia (hex) / 3 = Read Corrente / 4 = Read DCLink / 5 = Read Frequencia Hz / 6 = Status / 7 = Tensão de saida
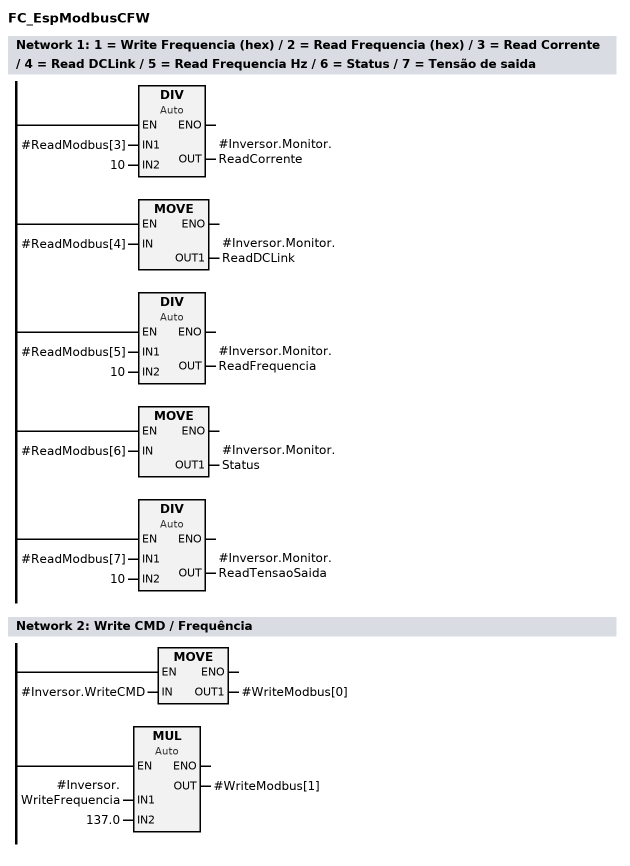
   RUNG wire#powerrail
      Div(in1 := #ReadModbus[3], in2 := 10, out => #Inversor.Monitor.ReadCorrente)
   END_RUNG
   RUNG wire#powerrail
      Move(in := #ReadModbus[4], out1 => #Inversor.Monitor.ReadDCLink)
   END_RUNG
   RUNG wire#powerrail
      Div(in1 := #ReadModbus[5], in2 := 10, out => #Inversor.Monitor.ReadFrequencia)
   END_RUNG
   RUNG wire#powerrail
      Move(in := #ReadModbus[6], out1 => #Inversor.Monitor.Status)
   END_RUNG
   RUNG wire#powerrail
      Div(in1 := #ReadModbus[7], in2 := 10, out => #Inversor.Monitor.ReadTensaoSaida)
   END_RUNG
   // the same network as SCL:
   #Inversor.Monitor.ReadCorrente := #ReadModbus[3] / 10;
   #Inversor.Monitor.ReadDCLink := #ReadModbus[4];
   #Inversor.Monitor.ReadFrequencia := #ReadModbus[5] / 10;
   #Inversor.Monitor.Status := #ReadModbus[6];
   #Inversor.Monitor.ReadTensaoSaida := #ReadModbus[7] / 10;
END_REGION

REGION Network 2: Write CMD / Frequência
   RUNG wire#powerrail
      Move(in := #Inversor.WriteCMD, out1 => #WriteModbus[0])
   END_RUNG
   RUNG wire#powerrail
      Mul(in1 := #Inversor.WriteFrequencia, in2 := 137.0, out => #WriteModbus[1])
   END_RUNG
   // the same network as SCL:
   #WriteModbus[0] := #Inversor.WriteCMD;
   #WriteModbus[1] := #Inversor.WriteFrequencia * 137.0;
END_REGION
END_FUNCTION

FUNCTION "FC_EspelhoModbusBal" : Void   // FC2, LAD
{ S7_Optimized_Access := 'TRUE' }
VERSION : 0.1
   VAR_IN_OUT
      ReadModbus : Array[0..6] of DInt;
      Balanca : "BalançaAlfa3101cs";
   END_VAR
BEGIN

REGION Network 1: Valor Negativo
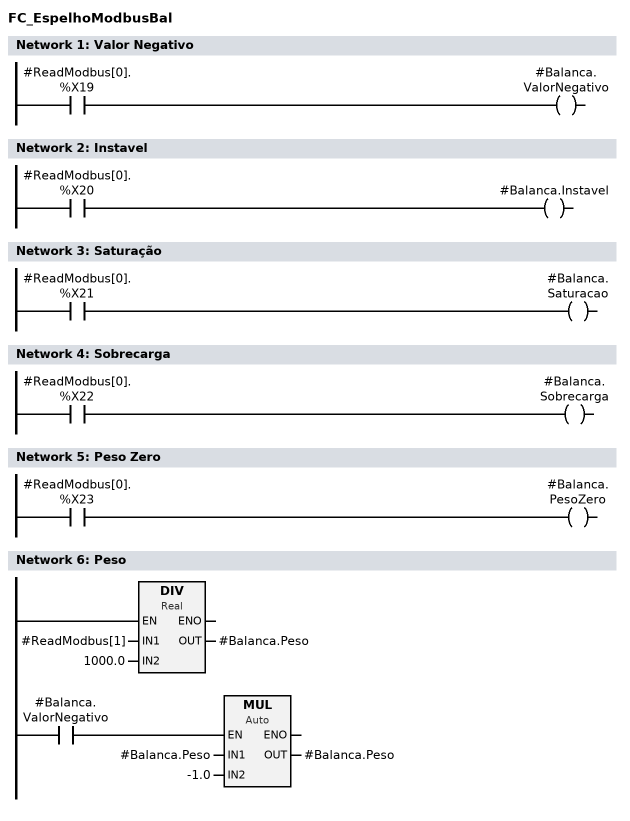
   RUNG wire#powerrail
      Contact( #ReadModbus[0].%X19 )
      Coil( #Balanca.ValorNegativo )
   END_RUNG
   // the same network as SCL:
   #Balanca.ValorNegativo := #ReadModbus[0].%X19;
END_REGION

REGION Network 2: Instavel
   RUNG wire#powerrail
      Contact( #ReadModbus[0].%X20 )
      Coil( #Balanca.Instavel )
   END_RUNG
   // the same network as SCL:
   #Balanca.Instavel := #ReadModbus[0].%X20;
END_REGION

REGION Network 3: Saturação
   RUNG wire#powerrail
      Contact( #ReadModbus[0].%X21 )
      Coil( #Balanca.Saturacao )
   END_RUNG
   // the same network as SCL:
   #Balanca.Saturacao := #ReadModbus[0].%X21;
END_REGION

REGION Network 4: Sobrecarga
   RUNG wire#powerrail
      Contact( #ReadModbus[0].%X22 )
      Coil( #Balanca.Sobrecarga )
   END_RUNG
   // the same network as SCL:
   #Balanca.Sobrecarga := #ReadModbus[0].%X22;
END_REGION

REGION Network 5: Peso Zero
   RUNG wire#powerrail
      Contact( #ReadModbus[0].%X23 )
      Coil( #Balanca.PesoZero )
   END_RUNG
   // the same network as SCL:
   #Balanca.PesoZero := #ReadModbus[0].%X23;
END_REGION

REGION Network 6: Peso
   RUNG wire#powerrail
      { S7_Templates := "SrcType := Real" } Div(in1 := #ReadModbus[1], in2 := 1000.0, out => #Balanca.Peso)
   END_RUNG
   RUNG wire#powerrail
      Contact( #Balanca.ValorNegativo )
      Mul(in1 := #Balanca.Peso, in2 := -1.0, out => #Balanca.Peso)
   END_RUNG
   // the same network as SCL:
   #Balanca.Peso := #ReadModbus[1] / 1000.0;
   IF #Balanca.ValorNegativo THEN #Balanca.Peso := #Balanca.Peso * (-1.0); END_IF;
END_REGION
END_FUNCTION

FUNCTION "FC_EspelhoModbusBal2711" : Void   // FC3, LAD
{ S7_Optimized_Access := 'TRUE' }
VERSION : 0.1
   VAR_IN_OUT
      ReadModbus : Array[0..8] of Int;
      WriteModBus : Array[0..8] of Word;
      Balanca : "BalançaAlfa3101cs";
   END_VAR
   VAR_TEMP
      DWord1 : DWord;
   END_VAR
BEGIN

REGION Network 1: Valor Negativo
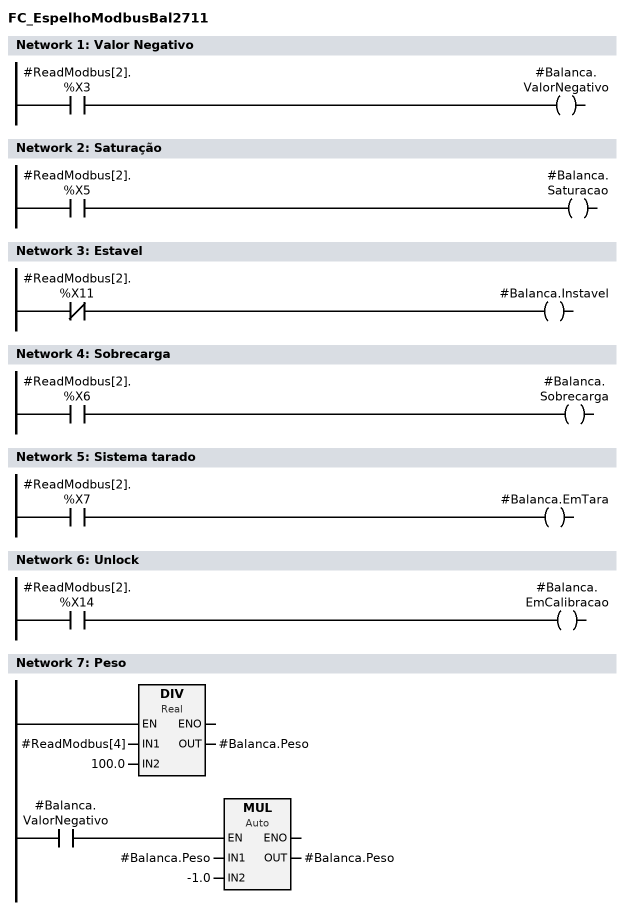
   RUNG wire#powerrail
      Contact( #ReadModbus[2].%X3 )
      Coil( #Balanca.ValorNegativo )
   END_RUNG
   // the same network as SCL:
   #Balanca.ValorNegativo := #ReadModbus[2].%X3;
END_REGION

REGION Network 2: Saturação
   RUNG wire#powerrail
      Contact( #ReadModbus[2].%X5 )
      Coil( #Balanca.Saturacao )
   END_RUNG
   // the same network as SCL:
   #Balanca.Saturacao := #ReadModbus[2].%X5;
END_REGION

REGION Network 3: Estavel
   RUNG wire#powerrail
      I_Contact( #ReadModbus[2].%X11 )
      Coil( #Balanca.Instavel )
   END_RUNG
   // the same network as SCL:
   #Balanca.Instavel := NOT #ReadModbus[2].%X11;
END_REGION

REGION Network 4: Sobrecarga
   RUNG wire#powerrail
      Contact( #ReadModbus[2].%X6 )
      Coil( #Balanca.Sobrecarga )
   END_RUNG
   // the same network as SCL:
   #Balanca.Sobrecarga := #ReadModbus[2].%X6;
END_REGION

REGION Network 5: Sistema tarado
   RUNG wire#powerrail
      Contact( #ReadModbus[2].%X7 )
      Coil( #Balanca.EmTara )
   END_RUNG
   // the same network as SCL:
   #Balanca.EmTara := #ReadModbus[2].%X7;
END_REGION

REGION Network 6: Unlock
   RUNG wire#powerrail
      Contact( #ReadModbus[2].%X14 )
      Coil( #Balanca.EmCalibracao )
   END_RUNG
   // the same network as SCL:
   #Balanca.EmCalibracao := #ReadModbus[2].%X14;
END_REGION

REGION Network 7: Peso
   RUNG wire#powerrail
      { S7_Templates := "SrcType := Real" } Div(in1 := #ReadModbus[4], in2 := 100.0, out => #Balanca.Peso)
   END_RUNG
   RUNG wire#powerrail
      Contact( #Balanca.ValorNegativo )
      Mul(in1 := #Balanca.Peso, in2 := -1.0, out => #Balanca.Peso)
   END_RUNG
   // the same network as SCL:
   #Balanca.Peso := #ReadModbus[4] / 100.0;
   IF #Balanca.ValorNegativo THEN #Balanca.Peso := #Balanca.Peso * (-1.0); END_IF;
END_REGION
END_FUNCTION

FUNCTION "FC_EspModbusFRECON" : Void   // FC4, LAD
{ S7_Optimized_Access := 'TRUE' }
VERSION : 0.1
   VAR_IN_OUT
      ReadModbus : Array[1..7] of Int;
      WriteFreq : Int;
      WriteCMD : Int;
      Inversor : "ModbusCFW";
   END_VAR
BEGIN

REGION Network 1: 3 = Read Corrente / 4 = Read DCLink / 5 = Read Frequencia Hz / 6 = Status / 7 = Tensão de saida
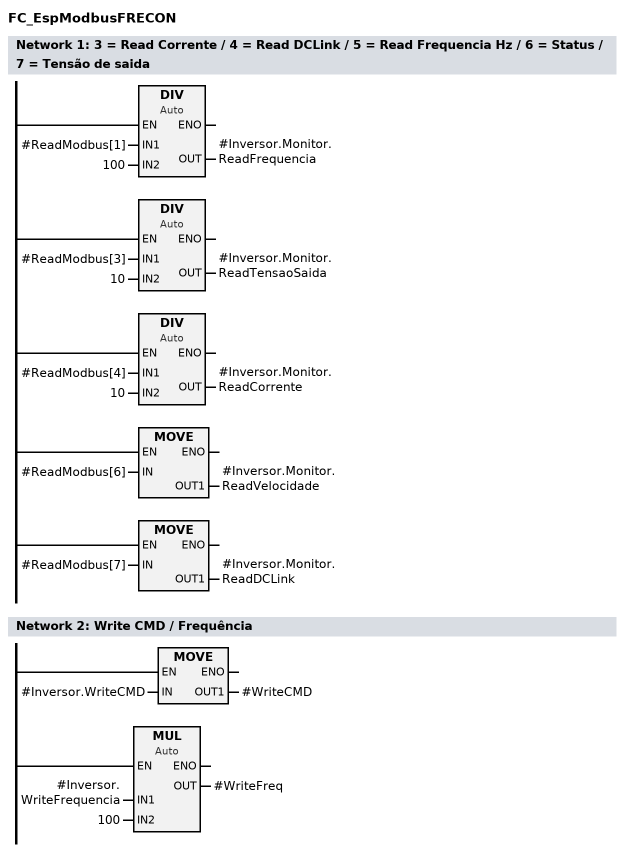
   RUNG wire#powerrail
      Div(in1 := #ReadModbus[1], in2 := 100, out => #Inversor.Monitor.ReadFrequencia)
   END_RUNG
   RUNG wire#powerrail
      Div(in1 := #ReadModbus[3], in2 := 10, out => #Inversor.Monitor.ReadTensaoSaida)
   END_RUNG
   RUNG wire#powerrail
      Div(in1 := #ReadModbus[4], in2 := 10, out => #Inversor.Monitor.ReadCorrente)
   END_RUNG
   RUNG wire#powerrail
      Move(in := #ReadModbus[6], out1 => #Inversor.Monitor.ReadVelocidade)
   END_RUNG
   RUNG wire#powerrail
      Move(in := #ReadModbus[7], out1 => #Inversor.Monitor.ReadDCLink)
   END_RUNG
   // the same network as SCL:
   #Inversor.Monitor.ReadFrequencia := #ReadModbus[1] / 100;
   #Inversor.Monitor.ReadTensaoSaida := #ReadModbus[3] / 10;
   #Inversor.Monitor.ReadCorrente := #ReadModbus[4] / 10;
   #Inversor.Monitor.ReadVelocidade := #ReadModbus[6];
   #Inversor.Monitor.ReadDCLink := #ReadModbus[7];
END_REGION

REGION Network 2: Write CMD / Frequência
   RUNG wire#powerrail
      Move(in := #Inversor.WriteCMD, out1 => #WriteCMD)
   END_RUNG
   RUNG wire#powerrail
      Mul(in1 := #Inversor.WriteFrequencia, in2 := 100, out => #WriteFreq)
   END_RUNG
   // the same network as SCL:
   #WriteCMD := #Inversor.WriteCMD;
   #WriteFreq := #Inversor.WriteFrequencia * 100;
END_REGION
END_FUNCTION

// ===== library types =====

// folder: 01_Blocks/Utilities

FUNCTION "LMQTT_ConvertToUtf8" : Void   // FC6, SCL
TITLE = LMQTT_ConvertToUtf8
{ S7_Optimized_Access := 'TRUE' }
AUTHOR : SIEMENS
FAMILY : LMQTT
VERSION : 1.0
// Function to convert a WCHAR to a UTF-8 conformant byte sequence
   VAR_INPUT
      character : WChar;   // Character that shall be converted to UTF-8
   END_VAR
   VAR_OUTPUT
      convertedUtf8 : DWord;   // UTF-8 conformant byte sequence. B0 stores first Byte, B1 second and B2 third Byte. B3 is not used
      bytesUsed : USInt;   // Amount of Bytes converted. Ranges from 1 to 3.
      error : Bool;   // TRUE: An error occurred during the execution of the FC
      status : Word;   // 16#0000 - 16#7FFF: Status of the FC, 16#8000 - 16#FFFF: Error identification
   END_VAR
   VAR_TEMP
      tempStatus : Word;   // temp value for output 'status'
      tempConvertedUtf8 : DWord;   // temp value for output 'convertedUtf8'
      tempBytesUsed : USInt;   // temp value for output 'bytesUsed'
      tempCharacter : WChar;   // temp value for input 'character'
   END_VAR
   // Ret_Val : No return for this FC - see error and status output
   VAR CONSTANT
      STATUS_NO_ERROR : Word := 16#0000;   // no error status
      STATUS_EXECUTION_FINISHED : Word := 16#0000;   // Execution finished without errors
      ERR_UNDEFINED : Word := 16#8000;   // Error due to an undefined case
      USINT_NULL : USInt := 0;   // Init value with 0
      DWORD_NULL : DWord := 16#0000_0000;   // Init value with 0
      EMPTY_WCHAR : WChar := WCHAR#' ';   // Empty WChar for comparison
      BELOW_7F : Word := 16#007F;   // Upper limit for character if only one Byte used
      BELOW_7FF : Word := 16#07FF;   // Upper limit for character if two Byte used
      BELOW_MAX_FFFF : Word := 16#FFFF;   // Upper limit for character if three Byte used
      BYTE_3F : Byte := 16#3F;   // Conversion Value
      BYTE_80 : Byte := 16#80;   // Conversion Value
      BYTE_C0 : Byte := 16#C0;   // Conversion Value
      BYTE_E0 : Byte := 16#E0;   // Conversion Value
      USINT_ONE : USInt := 1;   // Const Value to assign amount of bytes used
      USINT_TWO : USInt := 2;   // Const Value to assign amount of bytes used
      USINT_THREE : USInt := 3;   // Const Value to assign amount of bytes used
   END_VAR
BEGIN
   REGION BLOCK INFO HEADER
       //=============================================================================
       // SIEMENS AG
       // (c)Copyright 2020
       //-----------------------------------------------------------------------------
       // Library:       LMQTT
       // Tested with:   CPU 1516-3 PN/DP V2.8
       // Engineering:   TIA Portal V16
       // Restrictions:  --
       // Requirements:  --
       // Functionality: Converts a single WChar Character to a valid UTF-8 encoded byte sequence and saves this to a DWord.
       //                The amount of bytes saved is stored in bytesUsed Output.
       //-----------------------------------------------------------------------------
       // Change log table:
       // Version    Date         Expert in charge         Changes applied
       // 03.00.00   01.10.2020   Siemens Online Support   First released version
       //=============================================================================
   END_REGION

   REGION INITIALISATION  
       // Initialize functionality: reset of variables, diagnostics, etc.
       #tempConvertedUtf8 := #DWORD_NULL;
       #tempBytesUsed := #USINT_NULL;
       #tempStatus := #STATUS_NO_ERROR;
       //assign temp value from input:
        #tempCharacter := #character;

   END_REGION

   REGION PROGRAM LOGIC
       // Use this region for application specific code
       IF #tempCharacter = #EMPTY_WCHAR THEN
           //will be only 1 byte occupied
           #tempConvertedUtf8 := WCHAR_TO_DWORD(#tempCharacter);
           #tempBytesUsed := #USINT_ONE;
       ELSIF (WCHAR_TO_WORD(#tempCharacter) <= (#BELOW_7F)) THEN
           //will be only 1 byte occupied
           #tempConvertedUtf8 := WCHAR_TO_DWORD(#tempCharacter);
           #tempBytesUsed := #USINT_ONE;
       ELSIF (WCHAR_TO_WORD(#tempCharacter) <= (#BELOW_7FF)) THEN
           //will be 2 byte occupied
           #tempConvertedUtf8.%B1 := (WCHAR_TO_BYTE(#tempCharacter) AND #BYTE_3F) OR #BYTE_80;
           #tempConvertedUtf8.%B0 := WORD_TO_BYTE(SHR(IN := WCHAR_TO_WORD(#tempCharacter), N := 6)) OR #BYTE_C0;
           #tempBytesUsed := #USINT_TWO;
       ELSIF (WCHAR_TO_WORD(#tempCharacter) <= (#BELOW_MAX_FFFF)) THEN
           //will be 3 byte occupied
           #tempConvertedUtf8.%B2 := (WCHAR_TO_BYTE(#tempCharacter) AND #BYTE_3F) OR #BYTE_80;
           #tempConvertedUtf8.%B1 := (WORD_TO_BYTE(SHR(IN := WCHAR_TO_WORD(#tempCharacter), N := 6)) AND #BYTE_3F) OR #BYTE_80;
           #tempConvertedUtf8.%B0 := WORD_TO_BYTE(SHR(IN := WCHAR_TO_WORD(#tempCharacter), N := 12)) OR #BYTE_E0;
           #tempBytesUsed := #USINT_THREE;
       END_IF;
   END_REGION

   REGION OUTPUTS
       // Write application specific temp values to outputs
       #bytesUsed := #tempBytesUsed;
       #convertedUtf8 := #tempConvertedUtf8;
       // Write error and status
       #error := #tempStatus.%X15;
       #status := #tempStatus;
       // ENO mechanism is not used --> ENO := TRUE;
       ENO := TRUE;
   END_REGION
END_FUNCTION

// folder: Common

FUNCTION "IsIPAddress" : Bool   // FC1, SCL
TITLE = IsIPAddress
{ S7_Optimized_Access := 'TRUE' }
VERSION : 0.1
// Evaluates whether a given String contains a valid IP address
   VAR_INPUT
      address : String;   // Address to be evaluated
   END_VAR
   VAR_OUTPUT
      ipAddress : IP_V4;   // Parsed IP address if passed address is IP address
   END_VAR
   VAR_TEMP
      tempAddress : String;   // Passed address
      tempOctet : String;   // Current octet
      tempIndex : DInt;   // Index for loop
      tempPos : Int;   // Position of found separator
      tempNum : Int;   // Converted octet
      tempIp : IP_V4;   // Parsed IP address
   END_VAR
   // Ret_Val : Return value
   VAR CONSTANT
      MAX_VALUE : USInt := 255;   // Max. valid value of octet
      NUM_OCTETS : DInt := 4;   // Number of octets
      CHAR_ZERO : Char := '0';   // ASCII character '0'
   END_VAR
BEGIN
   REGION BLOCK INFO HEADER
     //===============================================================================
     // SIEMENS / (c)Copyright 2024
     //-------------------------------------------------------------------------------
     // Title:        IsIPAddress
     // Function:     Evaluates whether a given String contains a valid IP address
     // Library:      --
     // Author:       Siemens Industry Online Support
     // Tested with:  CPU 1515-2 PN V3.1
     // Engineering:  TIA Portal V17
     // Restrictions: --
     // Requirements: S7-1200 with firmware V4.4 or higher
     //               S7-1500 with firmware V2.0 or higher
     //-------------------------------------------------------------------------------
     // Change log table:
     // Version  | Date       | Expert in charge       | Changes applied
     //-------------------------------------------------------------------------------
     // 01.00.00 | 2024-02-12 | Online Support         | First released version
     //===============================================================================
   END_REGION

   #tempAddress := #address;
   #IsIPAddress := FALSE; // Will be overwritten if IP address is detected
   #ipAddress := #tempIp; // Zero output parameter

   FOR #tempIndex := 1 TO #NUM_OCTETS DO
     #tempPos := FIND(IN1 := #tempAddress, IN2 := '.'); // Find separator

     IF (#tempPos > 0 OR #tempIndex = #NUM_OCTETS) // Separator found with exception of last octet
       AND NOT (#tempPos > 0 AND #tempIndex = #NUM_OCTETS) // No separator found in last octet
       AND #tempPos <= 4 // 3  characters or less
     THEN
       IF #tempIndex < #NUM_OCTETS THEN // First three octets
         #tempOctet := LEFT(IN := #tempAddress, L := #tempPos - 1);
       ELSE// Last octet
         #tempOctet := #tempAddress;
       END_IF;

       STRG_VAL(IN := #tempOctet,
                FORMAT := 0,
                P := 1,
                OUT => #tempNum);

       IF #tempNum >= 0 AND #tempNum <= #MAX_VALUE // Within 0 and 255
         AND NOT (#tempNum = 0 AND #tempIndex = 1) // Not 0 in first octet
         AND NOT (#tempNum = 0 AND #tempOctet[1] <> #CHAR_ZERO) // Not 0 because of invalid character
       THEN
         #tempIp.ADDR[#tempIndex] := INT_TO_BYTE(#tempNum);
         #tempAddress := RIGHT(IN := #tempAddress, L := LEN(#tempAddress) - #tempPos); // Remove evaluated octet
       ELSE // Address is not IP address
         EXIT;
       END_IF;
     ELSE // Address is not IP address
       EXIT;
     END_IF;

     IF #tempIndex = #NUM_OCTETS THEN // End of loop reached, address is IP address
       #ipAddress := #tempIp;
       #IsIPAddress := true;
     END_IF;
   END_FOR;
END_FUNCTION

// folder: LMQTT

